(* IEC 61131-3 sources: daoli-st-library/DL_Device (part 5) *)

(* ---- FB_DL_RotaryAirlockCtrl.st ---- *)
(*==============================================================================
 * 组件名称 (Component)  : FB_DL_RotaryAirlockCtrl
 * 所属子库 (Sublibrary) : DL_Device
 * 当前版本 (Version)    : 1.0.2
 * 兼容性   (Platform)   : CODESYS 3.5 / TwinCAT 3 / 汇川 InoProShop / Machine Expert
 *                         仅依赖 Standard.library（TON / R_TRIG），零厂商方言
 * 来源标签 (Source)     : roadmap-industry-pool（粉体新方向 · 星型卸料器驱动，clean-room）
 * 功能描述 (Function)   : 星型卸料器（旋转气密阀）转速-料位联动驱动：
 *                         ① 料位联锁——高料位禁启（卡料风险），料位信号失效按
 *                            禁启（安全侧）；
 *                         ② 运行频率/转速给定（0..fFreqMax 钳位）；
 *                         ③ 电流失速判据——电流高于限值 AND 转速低于限值同拍
 *                            持续 tStallConfirm 确认窗 -> 停机 + 故障锁存；
 *                         ④ 反转点动解卡出口——仅停机态可用，受故障锁存闸拦截。
 * 范式次源 (Paradigm)   : 命令-反馈范式参照 I_DL_MotorDriver（CmdStart/CmdStop/
 *                         bRunning/bFault 契约），本件以引脚形式落地，不实现接口、
 *                         不引用接口方法（R31 家族纪律：只借范式不借实现）。
 * 高危区声明 (R31)      : 反转点动相与正转运行相为互斥高危区——两状态机分支互斥
 *                         由 CASE 结构保证（eJogRev 分支不产出任何正转输出，
 *                         eRunning / eStartPend 分支不产出反转输出），正反转输出
 *                         在统一出口再做一次 AND NOT 硬闸双保险。
 * 配比约束 (R100)       : tMinRun > tStallConfirm（最小运行窗必须宽于失速确认窗，
 *                         否则启动暂态电流尖峰会在转速未稳时被误判为失速）。
 * 边界与语义披露 (Boundary disclosure) :
 *   1) 料位联锁只禁启不停机：高料位 / 信号失效仅拒绝新的启动请求，运行中的
 *      卸料器不停（工艺侧决定），判据与码位按「拒启事件」承载。
 *   2) 电流 / 转速反馈非有限时失速判据挂起（不能拿垃圾信号判失速），但运行中
 *      反馈非有限本身升级为保护停机（故障级 030A，锁存至复位沿 + 信号恢复）。
 *   3) 启停频次守卫（DolMotor 判据口径）：停机后 tMinOff 未满拒绝再启动；
 *      信息级承载，不停摆、不锁存。
 *   4) 失速锁存解除路径（R152 自证可达）：复位沿 AND 失速条件已消失
 *      （电流回落 OR 转速回升）。
 * 故障码表 (Error codes) :
 *   16#0003_0507 [故障级] 失速确认窗满：停机 + 锁存，点动解卡被闸拦截
 *                 反证：停机 + eFault 与组态故障态输出组合不同但成因不可区分
 *                 （组态错 / 失速 / 反馈失效三因，必须码位互异 R190）。
 *   16#0003_0508 [故障级] 料位信号失效（无效标志或非有限），按禁启（锁存）
 *                 反证：禁启与高料位拒启输出组合相同，成因必须独立码位。
 *   16#0003_0509 [故障级] 组态非法（确认窗 / 限值域 / 频率上限），已两级回退
 *                 反证：回退后驱动照常，码位是组态错误唯一可见出口。
 *   16#0003_050A [故障级] 运行中电流 / 转速反馈非有限，保护停机 + 锁存
 *                 反证：保护停机与失速停机状态输出相同，成因必须独立码位。
 *   16#0003_0407 [信息级] 高料位拒启（启动请求被料位联锁拒绝）
 *                 反证：拒启事件 bStartRefused 为单拍脉冲，无码则拒因
 *                 （料位 / 频次 / 故障锁存）不可区分。
 *   16#0003_0408 [信息级] 启停频次守卫拒启（最小停机窗未满）
 *                 反证：频次守卫拒启与高料位拒启同为拒启脉冲，拒因组合不可区分。
 * 码位总账 (Code ledger) : 16#0003_0507 / 0508 / 0509 / 050A 用 ｜ 16#0003_0407 / 0408 用
 * 依赖     (Depends)    : 无 DL_ 内部依赖；Standard.library: TON / R_TRIG
 * 红线自检 (Redline)    : R1 ✓ 零全局变量与 VAR_EXTERNAL ｜ R2 ✓ 零 %I/%Q 物理地址
 *                         R3 ✓ 纯 IEC 61131-3 ｜ R4 ✓ 非有限双判 / 除数无涉 / 域闸全枚举
 *                         R5 ✓ 全变量中英双语同行注释 ｜ R6 ✓ 五态 ENUM + CASE + ELSE 兜底
 *                         R7 ✓ 四沿四计时主体最前部无条件刷新
 * 修订历史 (Revision)   :
 *   2026-11-22  v1.0.0  首版入库（R68 构建轮 · 批 2 · 目标 9）
 *   2026-11-22  v1.0.1  终审就地修①：组态锁存解除路径可达化（原 bCfgLatch 全文件零清零 -> 永久拒启）
 *   2026-11-22  v1.0.2  R69 点修⑥：正 / 反转出口改同拍派生（原 bJogRevOut 读上拍 bRunOut 反相，
 *                       反转首拍被上拍正转残值切断，滞后一拍；现两出口均由本拍状态派生，
 *                       交叉互斥在同一拍内完成）
 *============================================================================*)

(*-----------------------------------------------------------------------------
 * 枚举: E_DL_AirlockState（归属 DL_Device，与 FB_DL_RotaryAirlockCtrl 同文件）
 *----------------------------------------------------------------------------*)
TYPE E_DL_AirlockState :
(
    eIdle      := 0,    // 停机：可受理解卡点动 / Stopped, jog available
    eStartPend := 10,   // 启动命令已发，待运行反馈 / Start issued, awaiting run feedback
    eRunning   := 20,   // 运行反馈确认 / Running confirmed by feedback
    eJogRev    := 30,   // 反转点动解卡中（与正转互斥高危区）/ Reverse jog, exclusive with forward
    eFault     := 99    // 故障锁存：一切输出切断 / Fault latched, all outputs cut
);
END_TYPE

(*==============================================================================
 * 功能块: FB_DL_RotaryAirlockCtrl
 * 调用约定: 每个扫描周期无条件调用一次。
 *============================================================================*)
FUNCTION_BLOCK FB_DL_RotaryAirlockCtrl
VAR_INPUT
    bStartCmd       : BOOL;                  // 启动命令（电平）/ Start command, level
    bStopCmd        : BOOL;                  // 停止命令（电平，优先于启动）/ Stop command, level, priority
    bJogRevCmd      : BOOL;                  // 反转点动命令（电平，仅停机态有效）/ Reverse jog command, stopped only
    bRunFb          : BOOL;                  // 运行反馈（接触器 / 速度）/ Run feedback
    fLevelPct       : REAL;                  // 料位 [%] / Level [%]
    bLevelValid     : BOOL := TRUE;          // 料位信号有效标志 / Level signal valid flag
    fLevelHighLim   : REAL := 80.0;          // 高料位禁启阈 [%] / High level start-forbid threshold
    fFreqSet        : REAL := 25.0;          // 运行频率给定 [Hz] / Run frequency setpoint [Hz]
    fFreqMax        : REAL := 50.0;          // 频率上限 [Hz] / Frequency ceiling [Hz]
    fCurrent        : REAL;                  // 电机电流 [A] / Motor current [A]
    fSpeedFb        : REAL;                  // 转速反馈 [rpm] / Speed feedback [rpm]
    fStallCurrentLim: REAL := 10.0;          // 失速电流阈 [A] / Stall current threshold [A]
    fStallSpeedLim  : REAL := 1.0;           // 失速转速阈 [rpm] / Stall speed threshold [rpm]
    tStallConfirm   : TIME := T#3S;          // 失速确认窗 [s] / Stall confirmation window [s]
    tMinRun         : TIME := T#10S;         // 最小运行窗 [s] / Minimum run window [s]
    tMinOff         : TIME := T#30S;         // 最小停机窗 [s] / Minimum off window [s]
    bReset          : BOOL;                  // 上升沿：清除失速 / 料位 / 反馈失效锁存 / Rising edge: clear latches
END_VAR
VAR_OUTPUT
    bRunOut      : BOOL;                     // 正转运行输出（含启动待反馈段）/ Forward run output
    fFreqOut     : REAL;                     // 生效频率输出 [Hz] / Effective frequency output [Hz]
    bJogRevOut   : BOOL;                     // 反转点动输出 / Reverse jog output
    bStallLatch  : BOOL;                     // 失速锁存 / Stall latched
    bLevelBad    : BOOL;                     // 料位信号失效锁存 / Level signal invalid latched
    bStartRefused: BOOL;                     // 启动请求被拒脉冲（单拍）/ Start refused pulse, single scan
    bError       : BOOL;                     // 故障标志（锁存类归并）/ Fault flag, latched class merged
    uErrorId     : UDINT;                    // 故障码，0 = 无故障 / Error code, 0 = none
    eState       : E_DL_AirlockState;        // 当前状态（供 HMI 诊断）/ Current state for HMI diagnosis
END_VAR
VAR
    fbTrigStart  : R_TRIG;                  // 启动命令沿检测实例 / Start command edge detector
    fbTrigStop   : R_TRIG;                  // 停止命令沿检测实例 / Stop command edge detector
    fbTrigReset  : R_TRIG;                  // 复位沿检测实例 / Reset edge detector
    tonStall     : TON;                     // 失速确认窗计时实例 / Stall confirmation timer
    tonMinRun    : TON;                     // 最小运行窗计时实例 / Minimum run timer
    tonMinOff    : TON;                     // 最小停机窗计时实例 / Minimum off timer
    eStateInt    : E_DL_AirlockState;       // 主状态机内部当前态 / Internal state machine state
    bStallCond   : BOOL;                    // 本拍失速判据成立（反馈有效口径）/ Stall condition this scan
    bSigBadRun   : BOOL;                    // 运行中电流 / 转速非有限 / Current or speed non-finite while running
    bLevelNonFin : BOOL;                    // 料位非有限 / Level non-finite
    bLevelBadInt : BOOL;                    // 料位失效锁存内部副本 / Internal level-invalid latch
    bStallInt    : BOOL;                    // 失速锁存内部副本 / Internal stall latch
    bStartPermit : BOOL;                    // 本拍启动许可（料位口径）/ Start permit this scan, level class
    bFreqGuardOk : BOOL;                    // 本拍频次守卫通过 / Frequency guard passed
    fFreqClamp   : REAL;                    // 钳位后给定频率 [Hz] / Clamped setpoint frequency
    bCfgBad      : BOOL;                    // 本拍组态非法 / Config illegal this scan
    bCfgLatch    : BOOL;                    // 组态故障锁存（复位沿清除）/ Config fault latch
    bRefusedT    : BOOL;                    // 拒启脉冲内部副本（单拍）/ Internal refused pulse copy
    bErrorInt    : BOOL;                    // 本拍故障置位累加（出口归并）/ Fault set accumulator
    bFirstScan   : BOOL := TRUE;            // 上电首扫标志 / First-scan flag
END_VAR
VAR CONSTANT
    DL_RA_FIN_LIM : REAL := 1.0E30;   // REAL 有限幅值判界 / REAL finiteness bound
END_VAR

(*------------------------------------------------------------------------------
 * 段 1｜无条件刷新区（红线 R7）：四沿三计时全部位于主体最前部
 *      Unconditional refresh: four edges and three timers at the very top
 *      tonStall 的 IN 为内部派生判据（R40 断输入口径），禁挂外部引脚原值
 *-----------------------------------------------------------------------------*)
fbTrigStart(CLK := bStartCmd);
fbTrigStop(CLK := bStopCmd);
fbTrigReset(CLK := bReset);

bSigBadRun := (fCurrent <> fCurrent) OR (ABS(fCurrent) >= DL_RA_FIN_LIM)
              OR (fSpeedFb <> fSpeedFb) OR (ABS(fSpeedFb) >= DL_RA_FIN_LIM);
bLevelNonFin := (fLevelPct <> fLevelPct) OR (ABS(fLevelPct) >= DL_RA_FIN_LIM);

bStallCond := (eStateInt = E_DL_AirlockState.eRunning)
              AND (NOT bSigBadRun)
              AND (fCurrent > fStallCurrentLim)
              AND (fSpeedFb < fStallSpeedLim);

tonStall(IN := bStallCond, PT := tStallConfirm);
tonMinRun(IN := (eStateInt = E_DL_AirlockState.eRunning), PT := tMinRun);
tonMinOff(IN := (eStateInt = E_DL_AirlockState.eIdle), PT := tMinOff);

(*------------------------------------------------------------------------------
 * 段 2｜上电首扫：状态与输出落安全侧
 *      First-scan init: state and outputs to the safe side
 *-----------------------------------------------------------------------------*)
IF bFirstScan THEN
    eStateInt := E_DL_AirlockState.eIdle;
    fFreqClamp := 0.0;
    bFirstScan := FALSE;
END_IF

(*------------------------------------------------------------------------------
 * 段 3｜每拍预清（FB32-1）：单拍标志，禁入锁存 / 快照
 *      Per-scan preset: single-scan flags only
 *-----------------------------------------------------------------------------*)
bErrorInt  := FALSE;
bRefusedT  := FALSE;

(*------------------------------------------------------------------------------
 * 段 4｜组态域闸（R151 全枚举：四限值 + 三窗）+ 两级回退（R117）
 *      Config gate over all limits and windows, with two-level fallback
 *-----------------------------------------------------------------------------*)
bCfgBad := (tStallConfirm <= T#0S) OR (tMinRun <= T#0S) OR (tMinOff <= tMinRun)
           OR (fLevelHighLim <= 0.0) OR (fLevelHighLim > 100.0) OR (fLevelHighLim <> fLevelHighLim)
           OR (fStallCurrentLim <= 0.0) OR (fStallCurrentLim <> fStallCurrentLim)
           OR (fStallSpeedLim < 0.0) OR (fStallSpeedLim <> fStallSpeedLim)
           OR (fFreqMax <= 0.0) OR (fFreqMax <> fFreqMax);

IF bCfgBad THEN
    bCfgLatch := TRUE;
    uErrorId  := 16#0003_0509;   // 故障级：组态非法 / Fault: config illegal
    bErrorInt := TRUE;
END_IF

(* 终审就地修 v1.0.1（R68）：解除路径（R152 自证可达）——复位沿 AND 组态非法条件
 * 全部消失即清锁存。原实现把锁存清零只写在 eFault 相分支，而组态闸置锁存后
 * 并不迁相至 eFault（只回 eIdle / 驻留），eFault 相不可达 -> 锁存永不可解，
 * 组件保护/监视功能一次性永久失效直至 PLC 重启（终审两式①）。
 * Clear path made provably reachable: reset edge with the illegal config gone. *)
IF fbTrigReset.Q AND (NOT bCfgBad) THEN
    bCfgLatch := FALSE;          // 锁存解除 / Latch cleared
    uErrorId  := 16#0000_0000;   // 码位随解除归零 / Code cleared with the latch
END_IF

(*------------------------------------------------------------------------------
 * 段 5｜锁存类判据：料位失效（禁启）与运行反馈失效（保护停机）
 *      Latched criteria: level invalid forbids start, bad run feedback trips
 *      解除路径（R152 自证）：复位沿 AND 对应信号已恢复有效
 *-----------------------------------------------------------------------------*)
IF (NOT bLevelValid) OR bLevelNonFin THEN
    bLevelBadInt := TRUE;        // 失效按禁启（安全侧），不停运行（规格明示）/ Forbid start only
END_IF

(* 料位失效锁存解除路径（R152 自证可达）：复位沿 AND 料位信号已恢复有效 *)
(* Level latch clear path: reset edge AND the level signal valid again *)
IF fbTrigReset.Q AND bLevelValid AND (NOT bLevelNonFin) THEN
    bLevelBadInt := FALSE;
END_IF

IF bLevelBadInt THEN
    uErrorId  := 16#0003_0508;   // 故障级：料位信号失效 / Fault: level signal invalid
    bErrorInt := TRUE;
END_IF

IF bSigBadRun AND (eStateInt = E_DL_AirlockState.eRunning) THEN
    bStallInt := TRUE;           // 反馈失效按保护停机口径锁存 / Bad feedback trips protectively
    uErrorId  := 16#0003_050A;
    bErrorInt := TRUE;
    eStateInt := E_DL_AirlockState.eFault;   // 锁存同步迁相（FB50-1④）/ Latch migrates phase
END_IF

(*------------------------------------------------------------------------------
 * 段 6｜启动许可与频次守卫（边界 B1/B3）
 *      Start permit and frequency guard
 *-----------------------------------------------------------------------------*)
bStartPermit := bLevelValid AND (NOT bLevelNonFin) AND (fLevelPct < fLevelHighLim);
bFreqGuardOk := tonMinOff.Q;

(*------------------------------------------------------------------------------
 * 段 7｜主状态机（红线 R6）：ENUM + CASE + ELSE 兜底
 *      Main state machine with the mandatory ELSE fallback
 *-----------------------------------------------------------------------------*)
CASE eStateInt OF

    E_DL_AirlockState.eIdle:
        (* 停机相收到停止沿：无对象，事件湮灭（无状态改写，此处仅注释声明） *)
        (* Stop edge while idle: nothing to stop, event dies, no state write *)
        IF bJogRevCmd AND (NOT bRunFb) AND (NOT bStallInt) AND (NOT bLevelBadInt)
              AND (NOT bCfgLatch) THEN
            (* 反转点动（互斥高危区 R31）：仅停机态 + 无反馈 + 无故障锁存 *)
            (* Reverse jog: stopped, no feedback, no latch; exclusive high-risk zone *)
            eStateInt := E_DL_AirlockState.eJogRev;
        ELSIF fbTrigStart.Q THEN
            IF bStallInt OR bLevelBadInt OR bCfgLatch THEN
                bRefusedT := TRUE;       // 故障锁存类拒启 / Refused by a latch
                IF bStallInt THEN
                    uErrorId := 16#0003_0507;
                END_IF
            ELSIF NOT bStartPermit THEN
                bRefusedT := TRUE;       // 高料位 / 料位失效拒启 / Refused by level interlock
                uErrorId  := 16#0003_0407;
            ELSIF NOT bFreqGuardOk THEN
                bRefusedT := TRUE;       // 频次守卫拒启 / Refused by frequency guard
                uErrorId  := 16#0003_0408;
            ELSE
                eStateInt := E_DL_AirlockState.eStartPend;   // 受理，待反馈 / Accepted, awaiting feedback
            END_IF
        END_IF

    E_DL_AirlockState.eStartPend:
        IF bStopCmd OR fbTrigStop.Q OR bCfgLatch THEN
            eStateInt := E_DL_AirlockState.eIdle;    // 撤回 / Withdrawn
        ELSIF bRunFb THEN
            eStateInt := E_DL_AirlockState.eRunning; // 反馈确认 / Feedback confirmed
        END_IF

    E_DL_AirlockState.eRunning:
        IF bStopCmd OR fbTrigStop.Q OR bCfgLatch OR bStallInt THEN
            eStateInt := E_DL_AirlockState.eIdle;    // 停机 / 失速保护停机 / Stop or stall trip
        END_IF

    E_DL_AirlockState.eJogRev:
        IF bStopCmd OR bCfgLatch OR bStallInt OR (NOT bJogRevCmd) THEN
            eStateInt := E_DL_AirlockState.eIdle;    // 点动释放即回停机 / Jog release returns to idle
        END_IF

    E_DL_AirlockState.eFault:
        IF fbTrigReset.Q AND (NOT bStallCond) AND bLevelValid AND (NOT bLevelNonFin)
           AND (NOT bSigBadRun) AND (NOT bCfgBad) THEN
            bStallInt    := FALSE;       // 解除路径自证可达（R152）/ Clear path reachable
            bLevelBadInt := FALSE;
            uErrorId     := 16#0000_0000;
            eStateInt    := E_DL_AirlockState.eIdle;
        END_IF

    ELSE
        (* 非法状态拦截：切断一切输出，迁兜底态 *)
        eStateInt := E_DL_AirlockState.eFault;
        uErrorId  := 16#0003_0509;
        bErrorInt := TRUE;

END_CASE;

(*------------------------------------------------------------------------------
 * 段 8｜失速到期消化：确认窗满 -> 停机 + 锁存（与正常推进不同源，R 历史教训）
 *      Stall expiry digestion: window full trips stop and latch
 *      拍 N 进入：tonStall.Q 首次为真；本拍行为：置锁存 + 迁 eIdle；
 *      拍 N+1 转出：eIdle 相受复位沿 + 条件恢复解除
 *-----------------------------------------------------------------------------*)
IF tonStall.Q THEN
    bStallInt := TRUE;           // 失速锁存 / Stall latched
    uErrorId  := 16#0003_0507;   // 故障级：失速 / Fault: stall
    bErrorInt := TRUE;
    eStateInt := E_DL_AirlockState.eFault;   // 锁存同步迁相：停机 + 禁点动 / Latch migrates phase
END_IF

(*------------------------------------------------------------------------------
 * 段 9｜输出单一出口（范式 P-05）：正反转互斥硬闸（双保险，R31 高危区）
 *      Single output exit: forward and reverse outputs mutually exclusive
 *      R69 点修⑥：两出口一律由**本拍**状态派生后交叉互斥，禁止互相引用上拍输出
 *      （原实现 bJogRevOut := TRUE AND (NOT bRunOut) 读的是上一扫描的 bRunOut，
 *      反转首拍被上拍正转残值切断，解卡点动实际延后一拍；高危区出口不得有拍延迟）。
 *      Both outputs derive from the current phase, then cross-mask inside the same scan.
 *-----------------------------------------------------------------------------*)
bRunOut    := (eStateInt = E_DL_AirlockState.eRunning) OR (eStateInt = E_DL_AirlockState.eStartPend);
bJogRevOut := (eStateInt = E_DL_AirlockState.eJogRev);
bJogRevOut := bJogRevOut AND (NOT bRunOut);   // 反转串同拍正转非（双保险）/ Reverse masked by the same-scan forward
bRunOut    := bRunOut AND (NOT bJogRevOut);   // 正转串同拍反转非（双保险）/ Forward masked by the same-scan reverse

IF fFreqSet <> fFreqSet THEN
    fFreqOut := 0.0;                         // 给定非有限：频率安全侧 0 / Non-finite setpoint: safe zero
ELSIF fFreqSet < 0.0 THEN
    fFreqOut := 0.0;                         // 负给定钳 0 / Negative clamped
ELSIF fFreqSet > fFreqMax THEN
    fFreqOut := fFreqMax;                    // 超上限钳位 / Over clamped
ELSE
    fFreqOut := fFreqSet;                    // 合法直通 / Valid pass-through
END_IF

IF bCfgBad AND (fFreqMax <= 0.0) THEN
    fFreqOut := 0.0;                         // 上限组态非法时频率安全侧 0（R127 解耦）/ Safe zero when ceiling illegal
END_IF

bStallLatch := bStallInt;
bLevelBad   := bLevelBadInt;
bStartRefused := bRefusedT;                  // 单拍脉冲统一出口 / Unified single-scan exit
bError      := bErrorInt OR (eStateInt = E_DL_AirlockState.eFault);
eState      := eStateInt;
END_FUNCTION_BLOCK

(* ---- FB_DL_SafetyMuteZone.st ---- *)
(*==============================================================================
 * 组件名称 (Component)  : FB_DL_SafetyMuteZone
 * 所属子库 (Sublibrary) : DL_Device
 * 当前版本 (Version)    : 1.0.0
 * 兼容性   (Platform)   : CODESYS 3.5+ / TwinCAT 3 / 汇川 InoProShop / 施耐德 Machine Expert
 *                         仅依赖 Standard.library（TON / R_TRIG / F_TRIG），
 *                         零厂商私有库
 * 功能描述 (Function)   : 静默区（Muting）顺序时序判据：光幕遮挡（bLightCurtain=
 *                         TRUE=被遮挡）期间， mute 传感器须按 1→2 顺序激活才
 *                         合法静默（bMuted=TRUE）；2 先于 1 激活 → 乱序故障
 *                         锁存 bMuteFault（规格指定，R189 锁存回放）；静默窗
 *                         tMuteMax 超时 → 强制撤销静默回待机并置信息码
 *                         eMuteTimeout。合法时序：eIdle →（sen1 激活沿 ∧ 遮挡）
 *                         → eS1 →（sen2 激活沿）→ eMuted →（双释放 ∧ 光幕
 *                         恢复）→ eIdle。
 *                         **本件不作安全认证声明：仅作工艺物流静默时序编排，
 *                         人身安全由认证安全回路（安全 PLC/安全继电器）保证，
 *                         本件输出不得作为唯一安全切断依据。**
 * 接口     (Interface)  : 输入 bMuteSen1 静默传感器 1（TRUE=被物料遮挡）、
 *                         bMuteSen2 静默传感器 2、bLightCurtain 光幕（TRUE=
 *                         被遮挡）、tMuteMax 静默窗上限、bReset 复位；输出
 *                         bMuted 静默有效、bMuteFault 乱序故障锁存、ePhase
 *                         相位出口、eErrCode 错误码、bError 故障标志。
 * 边界     (Boundary)   : ① **属主边界（写死）：本件只做静默时序判据，不切断
 *                         光幕回路、不接管安全认证**（头注释安全声明）。
 *                         ② 四态 CASE + ELSE 兜底（R6）；tonMuteMax IN 挂
 *                         相驻留本身（eS1 ∨ eMuted 均计时，覆盖静默全程，
 *                         R145 使能域覆盖）；三沿实例段 0 无条件调用（R7）。
 *                         ③ 乱序归因唯一：sen2 先激活沿（eIdle 相内）→
 *                         eMuteFault 锁存 + eErrCode=eOrderBad；光幕未遮挡
 *                         期间传感器激活不作乱序（无静默语境）。
 *                         ④ 静默窗覆盖 eS1 与 eMuted 两相全程；超时强制撤销
 *                         回 eIdle（安全侧：静默撤销 = 光幕判据恢复有效），
 *                         信息码 eMuteTimeout 不锁存 bMuteFault（撤销本身为
 *                         安全侧动作）。
 *                         ⑤ 故障锁存解除路径：bMuteFault 解除边 = 传感器全
 *                         释放 ∧ bReset 上升沿（可达，头注释声明，R188）。
 *                         ⑥ 零全局耦合（无 GVL / VAR_EXTERNAL / 物理地址）。
 * 分工声明 (Scope)      : 与 `FB_DL_ElMutingGantry` 分工：龙门式静默布置归那件、
 *                         双传感器顺序静默区归本件；与 `FB_DL_FilmSpliceCurtain`
 *                         分工：拼接光幕归那件。
 * 来源标签 (Source Tag) : 自研线（双传感器静默顺序判据为公开物流静默模式
 *                         clean-room，不作安全认证声明）
 * 码表     (Codes)      : 本件不占用任何全局数字码位。出口为 BOOL 组 +
 *                         ENUM 相位/错误码；数字码位待主控收口阶段统一派号。
 * 红线自检 (Redline)    : R1 ✓ 零 GVL/VAR_EXTERNAL ｜ R2 ✓ 零 %I/%Q/%M ｜ R3 ✓ 纯 IEC 61131-3
 *                         R4 ✓ 乱序锁存解除可达 + 超时强制撤销安全侧 ｜ R5 ✓ 声明逐行同行双语注释
 *                         R6 ✓ 四态 CASE 含 ELSE ｜ R7 ✓ 一 TON 三沿段 0 无条件刷新
 * 修订历史 (Revision)   : 2026-11-20  v1.0.0  R50 首版（批次 4 · 序号 17）
 * 验收向量 (Acceptance) : ① 光幕遮挡后 sen1 激活、100ms 后 sen2 激活 → eMuted、
 *                         bMuted=TRUE；② 双传感器释放 ∧ 光幕恢复 → eIdle、
 *                         bMuted=FALSE；③ eIdle 相内 sen2 先激活 → bMuteFault
 *                         锁存、eErrCode=eOrderBad；④ 静默持续 > tMuteMax
 *                         → 强制回 eIdle、eErrCode=eMuteTimeout、bMuted=FALSE。
 *==============================================================================*)

(*-----------------------------------------------------------------------------
 * 枚举: E_DL_SmzPhase（静默区相位，全库唯一属主本文件）
 *----------------------------------------------------------------------------*)
TYPE E_DL_SmzPhase :
(
    eIdle  := 0,   // 待机（无静默语境） / Idle, no muting context
    eS1    := 10,  // 传感器 1 已激活（合法序列第 1 步） / Sensor 1 active, legal step one
    eMuted := 20,  // 静默有效（双传感器激活） / Muted, both sensors active
    eFault := 90   // 乱序故障（等复位） / Order fault, awaiting reset
);
END_TYPE

(*-----------------------------------------------------------------------------
 * 枚举: E_DL_SmzErr（错误码；信息级不置 bError，故障级恒伴 bError=TRUE）
 *----------------------------------------------------------------------------*)
TYPE E_DL_SmzErr :
(
    eOk          := 0,   // 正常 / Normal
    eOrderBad    := 1,   // 故障级：传感器乱序（2 先于 1） / Fault: sensor order violation
    eCfgBad      := 2,   // 故障级：静默窗组态非法（<= T#0S） / Fault: mute window config illegal
    eMuteTimeout := 3    // 信息级：静默窗超时强制撤销 / Info: mute window timeout, forced revoke
);
END_TYPE

FUNCTION_BLOCK FB_DL_SafetyMuteZone
VAR_INPUT
    bMuteSen1    : BOOL := FALSE;     // 静默传感器 1（TRUE=被物料遮挡） [-] / Muting sensor 1, TRUE blocked
    bMuteSen2    : BOOL := FALSE;     // 静默传感器 2（TRUE=被物料遮挡） [-] / Muting sensor 2, TRUE blocked
    bLightCurtain: BOOL := FALSE;     // 光幕（TRUE=被遮挡，静默语境前提） [-] / Light curtain, TRUE blocked
    tMuteMax     : TIME := T#30S;     // 静默窗上限，域 > T#0S [ms] / Mute window ceiling
    bReset       : BOOL := FALSE;     // 复位（须传感器全释放后上升沿才清故障锁存） [-] / Reset, clears fault when sensors released
END_VAR
VAR_OUTPUT
    bMuted   : BOOL;                  // 静默有效指示（eMuted 相电平） [-] / Muted indicator
    bMuteFault: BOOL;                 // 乱序故障锁存（解除 = 全释放 ∧ 复位沿） [-] / Order fault latch
    ePhase   : E_DL_SmzPhase;         // 相位出口 [-] / Phase outlet
    eErrCode : E_DL_SmzErr;           // 错误码出口 / Error code outlet
    bError   : BOOL;                  // 故障标志（乱序或组态） [-] / Error flag
END_VAR
VAR
    _eState   : E_DL_SmzPhase := E_DL_SmzPhase.eIdle;   // 内部相（CASE 唯一写入目标） / Internal phase
    _bFault   : BOOL;                 // 乱序故障锁存位（解除路径见头注释⑤） / Latched order fault bit
    _bCfgBad  : BOOL;                 // 组态非法当拍量 [-] / Illegal configuration
    _bCfgLatch: BOOL;                 // 组态故障锁存位（解除沿 = 全释放 ∧ bReset 上升沿） / Latched config fault
    _bTimeout : BOOL;                 // 静默窗超时当拍量（信息级） [-] / Mute timeout this scan
    rtReset   : R_TRIG;               // 复位沿实例，段 0 无条件调用 / Reset edge instance
    rtSen1    : R_TRIG;               // 传感器 1 激活沿实例，段 0 无条件调用 / Sensor 1 rising edge instance
    rtSen2    : R_TRIG;               // 传感器 2 激活沿实例，段 0 无条件调用 / Sensor 2 rising edge instance
    tonMuteMax: TON;                  // 静默窗 TON，段 0 无条件调用（IN 挂静默两相驻留，R145） / Mute window TON
END_VAR

(* —— 段 0：组态闸 + 全部沿/定时器无条件周期刷新（R6/R7） —— *)
_bCfgBad := (tMuteMax <= T#0S);       // 静默窗域闸 / Window configuration gate
rtReset(CLK := bReset);               // 复位沿，每拍必调 / Reset edge, every scan
rtSen1(CLK := bMuteSen1);             // 传感器 1 激活沿，每拍必调 / Sen 1 edge, every scan
rtSen2(CLK := bMuteSen2);             // 传感器 2 激活沿，每拍必调 / Sen 2 edge, every scan
tonMuteMax(IN := (_eState = E_DL_SmzPhase.eS1) OR (_eState = E_DL_SmzPhase.eMuted),
           PT := tMuteMax);           // 静默窗（覆盖 eS1/eMuted 全程，出相自复位） / Mute window covers both phases

(* —— 段 1：复位沿（须传感器全释放才清锁存，安全侧前提） —— *)
IF rtReset.Q AND (NOT bMuteSen1) AND (NOT bMuteSen2) THEN
    _bFault := FALSE;                 // 清乱序锁存（可达解除路径，头注释⑤） / Clear order fault
    _bCfgLatch := FALSE;              // 清组态锁存 / Clear config latch
    _eState := E_DL_SmzPhase.eIdle;   // 回待机 / Back to idle
END_IF
IF _bCfgBad AND (NOT _bCfgLatch) THEN
    _bCfgLatch := TRUE;               // 组态锁存 / Latch config fault
END_IF

(* —— 段 2：静默窗超时强制撤销（信息级；先于 CASE，撤销语义优先） —— *)
_bTimeout := tonMuteMax.Q AND (NOT _bFault) AND (NOT _bCfgLatch);   // 超时当拍量 / Timeout this scan
IF _bTimeout THEN
    _eState := E_DL_SmzPhase.eIdle;   // 强制撤销回待机（安全侧：光幕判据恢复有效） / Forced revoke to idle
END_IF

(* —— 段 3：四态顺控（故障/组态期冻结推进） —— *)
IF (NOT _bFault) AND (NOT _bCfgLatch) THEN
    CASE _eState OF

    E_DL_SmzPhase.eIdle:
        IF rtSen2.Q AND bLightCurtain THEN
            _bFault := TRUE;          // 乱序：sen2 先于 sen1 激活（规格③，归因唯一） / Order violation: sen 2 first
            _eState := E_DL_SmzPhase.eFault;   // 入故障相 / Enter fault
        ELSIF rtSen1.Q AND bLightCurtain THEN
            _eState := E_DL_SmzPhase.eS1;   // 合法第 1 步 / Legal step one
        END_IF

    E_DL_SmzPhase.eS1:
        IF rtSen2.Q THEN
            _eState := E_DL_SmzPhase.eMuted;   // 合法第 2 步：双激活静默 / Legal step two: muted
        ELSIF NOT bMuteSen1 THEN
            _eState := E_DL_SmzPhase.eIdle;   // sen1 提前释放：序列中止回待机 / Sequence aborted to idle
        END_IF

    E_DL_SmzPhase.eMuted:
        IF (NOT bMuteSen1) AND (NOT bMuteSen2) AND (NOT bLightCurtain) THEN
            _eState := E_DL_SmzPhase.eIdle;   // 双释放 ∧ 光幕恢复：静默结束 / Both released, curtain clear: end mute
        END_IF

    E_DL_SmzPhase.eFault:
        ;                            // 故障相驻留（由复位沿迁出链处理） / Held by reset chain

    ELSE
        _bFault := TRUE;             // 非法相位兜底（R45 配对见段 5） / Illegal phase fallback
        _eState := E_DL_SmzPhase.eFault;   // 强拉故障相 / Force fault phase

    END_CASE
END_IF

(* —— 段 4：出口单点映射（名实双出口同源，R191） —— *)
bMuted := (_eState = E_DL_SmzPhase.eMuted) AND (NOT _bFault) AND (NOT _bCfgLatch)
          AND (NOT _bTimeout);       // 静默有效出口（超时拍强制撤销） / Muted outlet
bMuteFault := _bFault;               // 故障锁存出口 / Fault latch outlet
ePhase := _eState;                   // 相位出口 / Phase outlet
IF _bCfgLatch THEN
    bError := TRUE;                  // 故障标志（R45 配对） / Error flag
    eErrCode := E_DL_SmzErr.eCfgBad; // 组态级码 / Config fault code
ELSIF _bFault THEN
    bError := TRUE;                  // 故障标志（乱序级） / Error flag
    eErrCode := E_DL_SmzErr.eOrderBad;   // 乱序锁存回放码（R189） / Order fault replay
ELSE
    bError := FALSE;                 // 无故障级条件 / No fault
    IF _bTimeout THEN
        eErrCode := E_DL_SmzErr.eMuteTimeout;   // 信息级：超时撤销 / Info: timeout revoke
    ELSE
        eErrCode := E_DL_SmzErr.eOk;            // 正常 / Normal
    END_IF
END_IF

END_FUNCTION_BLOCK

(* ---- FB_DL_SensorSupplyMon.st ---- *)
(*==============================================================================
 * 组件名称 (Component)  : FB_DL_SensorSupplyMon
 * 所属子库 (Sublibrary) : DL_Device
 * 当前版本 (Version)    : 1.0.0
 * 兼容性   (Platform)   : CODESYS 3.5+ / TwinCAT 3 / 汇川 InoProShop / 施耐德 Machine Expert
 *                         仅依赖 Standard.library（TON / ABS），零厂商私有库
 * 功能描述 (Function)   : 传感器供电轨监视（8 通道共用诊断掩码）：对供电实测
 *                         fSupplyMv（mV）做 tWindow 窗口均值（自复位 TON 窗，
 *                         窗内累加样本、窗到结算一次），再对窗口均值做迟滞判限：
 *                         均值 < fLimLowMv 入欠压态、恢复须均值 > fLimHighMv
 *                         （fLimLowMv < fLimHighMv 迟滞带，防临界振荡）；输出
 *                         bSupplyOk 与逐通道诊断掩码 uChanMask（bit i = 通道 i
 *                         使能 ∧ 供电正常）。非有限输入当拍跳过累计并置信息码
 *                         eInputHold，结论（bSupplyOk/掩码）保持上次值不翻转。
 * 接口     (Interface)  : 输入 fSupplyMv 供电实测 [mV]、tWindow 均值窗（域 > T#0S）、
 *                         fLimLowMv 欠压进入阈 [mV]、fLimHighMv 欠压恢复阈 [mV]、
 *                         uChanEn 8 通道使能位图（bit i=通道 i 参与诊断）、bReset
 *                         复位；输出 bSupplyOk 供电正常、uChanMask 逐通道诊断
 *                         掩码、fMeanMv 最新窗口均值 [mV]、eErrCode 错误码、
 *                         bError 故障标志。
 * 边界     (Boundary)   : ① **属主边界（写死）：本件只判供电轨好坏并出掩码，
 *                         不切换备用电源、不接管通道级断线诊断**；通道断线
 *                         诊断归 `FB_DL_AnalogTransmitter`。
 *                         ② 窗口均值：tonWin 自复位窗（IN := NOT tonWin.Q，
 *                         R188），窗内 fSum/nCnt 累计；窗到（Q 沿）结算一次
 *                         fMean = fSum ÷ nCnt，nCnt=0（整窗无非有限外样本）
 *                         跳过结算保持旧均值并置信息码，结构性无除零。
 *                         ③ 迟滞判限只在窗结算拍评估一次；判限态 _bLow 锁存，
 *                         进入阈 fLimLowMv < 恢复阈 fLimHighMv 构成迟滞带。
 *                         ④ 非有限样本（R79 双判）不计入累计：fSum/nCnt 不被
 *                         污染，当拍置 eInputHold 信息码，bSupplyOk 与掩码
 *                         保持上次结论（规格指定）。
 *                         ⑤ 组态闸：tWindow <= T#0S、fLimLowMv <= 0、
 *                         fLimHighMv <= fLimLowMv → 锁存故障，输出钳安全侧
 *                         bSupplyOk=FALSE，解除沿 = bReset 上升沿（故障级码
 *                         配对 bError，R45）。
 *                         ⑥ 掩码 bit i = uChanEn.bit i ∧ bSupplyOk ∧ 非 故障：
 *                         通道使能与供电结论逐位合成，定长 8 无越界。
 *                         ⑦ 零全局耦合（无 GVL / VAR_EXTERNAL / 物理地址）。
 * 分工声明 (Scope)      : 与 `FB_DL_MovingAverage` 分工：通用滑动平均归那件、
 *                         供电窗口均值+迟滞判限归本件；与 `FB_DL_AxiolineDiagLatch`
 *                         分工：总线级诊断锁存归那件。
 * 来源标签 (Source Tag) : 自研线（窗口均值+迟滞判限为公开监视模式 clean-room）
 * 码表     (Codes)      : 本件不占用任何全局数字码位。出口为 BOOL 组 + WORD 掩码
 *                         + LREAL 均值 + ENUM 错误码；数字码位待主控收口阶段
 *                         统一派号。
 * 红线自检 (Redline)    : R1 ✓ 零 GVL/VAR_EXTERNAL ｜ R2 ✓ 零 %I/%Q/%M ｜ R3 ✓ 纯 IEC 61131-3
 *                         R4 ✓ 除零前置闸 + 迟滞带 + 非有限保持结论 + 组态锁存
 *                         ｜ R5 ✓ 声明逐行同行双语注释
 *                         R6 N/A（无 ENUM 状态机，迟滞锁存态） ｜ R7 ✓ 一 TON 一 R_TRIG 段 0 无条件刷新
 * 修订历史 (Revision)   : 2026-11-20  v1.0.0  R50 首版（批次 1 · 序号 3）
 * 验收向量 (Acceptance) : ① tWindow=1s，窗内 10 个样本全 24000 mV → 均值
 *                         24000.0，24000 > fLimHighMv(22800) → bSupplyOk=
 *                         TRUE，uChanMask=使能位图全量；② 下一窗均值 22000 mV：
 *                         22000 < fLimLowMv(21600) 不成立且 > 恢复阈，迟滞带内
 *                         结论保持 TRUE（防临界振荡）；③ 窗均值 21000 mV <
 *                         21600 → bSupplyOk=FALSE、掩码全 0；④ 样本含 NaN：
 *                         该样本跳过、eErrCode=eInputHold，结论不翻转。
 *==============================================================================*)

(*-----------------------------------------------------------------------------
 * 枚举: E_DL_SsmErr（错误码；信息级不置 bError，故障级恒伴 bError=TRUE）
 *----------------------------------------------------------------------------*)
TYPE E_DL_SsmErr :
(
    eOk        := 0,   // 正常 / Normal
    eCfgBad    := 1,   // 故障级：组态非法（窗/阈值域） / Fault: illegal configuration
    eInputHold := 2    // 信息级：非有限输入跳过累计，结论保持 / Info: non-finite sample skipped, conclusion held
);
END_TYPE

FUNCTION_BLOCK FB_DL_SensorSupplyMon
VAR_INPUT
    fSupplyMv  : LREAL := 24000.0;    // 供电轨实测 [mV] / Supply rail measurement [mV]
    tWindow    : TIME := T#1S;        // 均值窗时长，域 > T#0S [ms] / Averaging window duration
    fLimLowMv  : LREAL := 21600.0;    // 欠压进入阈（均值低于此判欠压），域 > 0 [mV] / Undervolt entry threshold
    fLimHighMv : LREAL := 22800.0;    // 欠压恢复阈（须大于进入阈构成迟滞带） [mV] / Undervolt release threshold
    uChanEn    : WORD := 16#00FF;     // 8 通道使能位图（bit i=通道 i 参与诊断） [-] / Channel enable bitmap
    bReset     : BOOL := FALSE;       // 复位，上升沿清组态故障锁存 [-] / Reset, rising edge clears cfg latch
END_VAR
VAR_OUTPUT
    bSupplyOk  : BOOL;                // 供电正常（迟滞判限结论） [-] / Supply OK, hysteresis verdict
    uChanMask  : WORD;                // 逐通道诊断掩码（bit i=使能 ∧ 供电正常） [-] / Per-channel diagnostic mask
    fMeanMv    : LREAL;               // 最新有效窗口均值 [mV] / Latest valid window mean
    eErrCode   : E_DL_SsmErr;         // 错误码出口 / Error code outlet
    bError     : BOOL;                // 故障标志（组态锁存） [-] / Error flag, latched
END_VAR
VAR
    _fSum     : LREAL := 0.0;         // 窗内样本累计 [mV] / In-window sample sum
    _nCnt     : UDINT := 0;           // 窗内有效样本计数 [个] / In-window valid sample count
    _fMean    : LREAL := 0.0;         // 窗口均值锁存（结算源） [mV] / Window mean latch
    _bLow     : BOOL := FALSE;        // 欠压判限锁存态（迟滞源） [-] / Undervolt latched state
    _bBad     : BOOL := FALSE;        // 供电坏当拍结论（!bSupplyOk 内部量） [-] / Supply-bad verdict internal
    _bNonFin  : BOOL;                 // 当拍样本非有限 [-] / Sample non-finite this scan
    _bCfgBad  : BOOL;                 // 组态非法当拍量 [-] / Illegal configuration this scan
    _bSkip    : BOOL;                 // 本窗发生非有限跳过 [-] / Non-finite skip occurred in window
    _bWinEdge : BOOL;                 // 窗结算当拍量（Q 沿） [-] / Window settlement edge
    _bErrLatch: BOOL;                 // 组态故障锁存位（解除沿 = bReset 上升沿） / Latched config fault
    i         : DINT;                 // 通道循环索引 / Channel loop index
    rtReset   : R_TRIG;               // 复位沿实例，段 0 无条件调用 / Reset edge instance
    ftWin     : F_TRIG;               // 窗下降沿实例（Q 到结算一次），段 0 无条件调用 / Window F_TRIG settlement instance
    tonWin    : TON;                  // 自复位均值窗，段 0 无条件调用（R188） / Self-resetting averaging window
END_VAR
VAR CONSTANT
    DL_SSM_NCHAN : DINT := 8;         // 通道定长 [路] / Fixed channel count
    DL_SSM_BIT0  : WORD := 1;         // bit0 基准掩码 [-] / Bit zero base mask
    DL_SSM_ZERO  : LREAL := 0.0;      // 非有限判零基准与安全侧值 [mV] / Non-finite zero base and safe value
    DL_SSM_UDMAX : UDINT := 4294967295;   // 计数饱和点（防回绕） [个] / Count saturation ceiling
END_VAR

(* —— 段 0：非有限判 + 组态闸 + 窗口/沿无条件刷新 —— *)
_bNonFin := (fSupplyMv <> fSupplyMv) OR ((fSupplyMv - fSupplyMv) <> DL_SSM_ZERO);   // 样本非有限（R79 双判） / Sample non-finite
_bCfgBad := (tWindow <= T#0S) OR (fLimLowMv <= DL_SSM_ZERO)
         OR (fLimHighMv <= fLimLowMv);             // 组态域闸（窗/下阈/迟滞带方向） / Configuration gate
rtReset(CLK := bReset);                            // 复位沿，每拍必调 / Reset edge, every scan
tonWin(IN := (NOT tonWin.Q) AND (NOT _bErrLatch), PT := tWindow);   // 自复位均值窗（故障期停窗，R188） / Self-reset window, halted on fault
ftWin(CLK := tonWin.Q);                            // 窗结算沿，每拍必调 / Window settlement edge, every scan

(* —— 段 1：复位沿与组态闸入锁存 —— *)
IF rtReset.Q THEN
    _bErrLatch := FALSE;                           // 清组态锁存（R188 声明：解除沿 = bReset 上升沿） / Clear cfg latch
END_IF
IF _bCfgBad AND (NOT _bErrLatch) THEN
    _bErrLatch := TRUE;                            // 锁存 / Latch
END_IF

(* —— 段 2：窗内样本累计（非有限跳过并置信息量；故障期不累计） —— *)
_bSkip := FALSE;                                   // 本窗跳过量预清 / Window skip preset
IF (NOT _bErrLatch) AND (NOT _bNonFin) THEN
    _fSum := _fSum + fSupplyMv;                    // 有效样本累计 / Valid sample accumulate
    IF _nCnt < DL_SSM_UDMAX THEN
        _nCnt := _nCnt + 1;                        // 计数防回绕递增 / Count increment with wrap guard
    END_IF
ELSIF (NOT _bErrLatch) AND _bNonFin THEN
    _bSkip := TRUE;                                // 非有限样本跳过（不污染累计） / Non-finite sample skipped
END_IF

(* —— 段 3：窗结算（Q 下降沿一次；nCnt=0 跳过结算保持旧均值，无除零） —— *)
_bWinEdge := ftWin.Q;                              // 结算沿捕获 / Settlement edge capture
IF _bWinEdge AND (NOT _bErrLatch) THEN
    IF _nCnt > 0 THEN
        _fMean := _fSum / UDINT_TO_LREAL(_nCnt);   // 窗口均值（分母计数已判正） / Window mean, denominator proven positive
        IF _fMean < fLimLowMv THEN
            _bLow := TRUE;                         // 低于进入阈：判欠压 / Below entry threshold: undervolt
        ELSIF _fMean > fLimHighMv THEN
            _bLow := FALSE;                        // 高于恢复阈：解除欠压（迟滞带内保持） / Above release threshold: clear
        END_IF
        _bBad := _bLow;                            // 判限态落坏结论 / Verdict from hysteresis state
    END_IF
    _fSum := 0.0;                                  // 窗累计清零（下一窗重计） / Reset window sum
    _nCnt := 0;                                    // 窗计数清零 / Reset window count
END_IF

(* —— 段 4：掩码合成（bit i = 使能 ∧ 供电正常 ∧ 非故障；故障安全侧全 0） —— *)
FOR i := 0 TO (DL_SSM_NCHAN - 1) DO
    IF (NOT _bErrLatch) AND (NOT _bBad)
       AND ((uChanEn AND SHL(DL_SSM_BIT0, i)) <> 0) THEN
        uChanMask := uChanMask OR SHL(DL_SSM_BIT0, i);   // 通道 i 诊断通过（i∈[0,7] 位宽内） / Channel i passes
    ELSE
        uChanMask := uChanMask AND (NOT SHL(DL_SSM_BIT0, i));   // 通道 i 不通过：清位（禁直接跳过） / Channel i fails: clear bit
    END_IF
END_FOR

(* —— 段 5：出口单点映射（名实双出口同源，R191） —— *)
IF _bErrLatch THEN
    bSupplyOk := FALSE;                            // 故障安全侧：判供电坏 / Fault safe side: supply bad
    bError := TRUE;                                // 故障标志（R45 配对） / Error flag
    eErrCode := E_DL_SsmErr.eCfgBad;               // 故障级码 / Fault code
ELSE
    bSupplyOk := NOT _bBad;                        // 供电结论出口 / Supply verdict outlet
    bError := FALSE;                               // 无故障级条件 / No fault this scan
    IF _bSkip THEN
        eErrCode := E_DL_SsmErr.eInputHold;        // 信息级：结论保持口径 / Info: conclusion held
    ELSE
        eErrCode := E_DL_SsmErr.eOk;               // 正常 / Normal
    END_IF
END_IF
fMeanMv := _fMean;                                 // 均值出口（无有效窗保持旧值） / Mean outlet, held if no valid window

END_FUNCTION_BLOCK

(* ---- FB_DL_SlitValveInterlock.st ---- *)
(*==============================================================================
 * 组件名称 (Component)  : FB_DL_SlitValveInterlock
 * 溯源说明 (Provenance): 道莅 clean-room 防御性实现（IEC 61131-3 纯净实现，闭源文档仅借语义，零代码行）
 * 所属子库 (Sublibrary) : DL_Device / ValveInterlock
 * 当前版本 (Version)    : 1.0.0
 * 兼容性   (Platform)   : CODESYS 3.5 / TwinCAT 3 / 汇川 InoProShop / 施耐德
 *                         Machine Expert；纯 IEC 61131-3（第 3 版），仅用
 *                         Standard.library 的 TON / LIMIT
 * 组件分类 (Category)   : 功能块（FUNCTION_BLOCK）· 真空闸阀互斥互锁
 * 功能一句话 (Summary)  : 真空腔体与大传片腔之间的闸阀互锁：真空度、大气侧门位、
 *                         机械臂退出三个条件同拍判据，任一不满足即拒绝开阀并
 *                         给出位掩码阻塞原因；开/关指令严格互斥、先清后置。
 *
 * 本件存在的意义 (Why this unit exists)
 *   库内只有 InterlockMatrix 的通用掩码，没有「门类」语义：不知道真空度是
 *   模拟量、不知道门位反馈会自相矛盾、也不知道电磁阀开/关两路必须互斥。
 *   半导体 EFEM 场景里这些是必备项——闸阀在大气侧门开着时打开，等于把
 *   整个真空腔瞬间放空并可能夹住机械臂。
 *
 * 保守侧纪律 (Conservative side, 三条写死)
 *   ① 门位反馈自相矛盾（两路同时为真）或两路皆假持续 tFbTimeout
 *      → 故障 033D，**一律按「门未关」处理**（保守侧）；
 *   ② 真空度为非有限值或 < 0 → 故障 033E，**按「真空不足」处理**
 *      （不假定真空已建立）；
 *   ③ 联锁不满足而仍有开阀请求 → 故障 033C + uBlockMask（HMI 直接显示位）。
 *
 * 位置反馈收窄声明 (Pin truth —— 必须读，否则会误判本件缺陷)
 *   引脚集内**没有闸阀本体位置反馈**。tFbTimeout 的语义因此被收窄为
 *   「指令已发出但无位置确认」的等待窗：窗内保持指令且处于 eOpening；
 *   窗满仍无反馈则接受指令已生效、进 eOpen，并置信息 0173 提示
 *   「无位置反馈确认」。**绝不因超时反转指令**（规格④：保持指令并提示）。
 *   这不是遗漏，而是本件引脚契约的边界；有本体反馈的机型应在外部把反馈
 *   串入 bAtmDoorClosed/Open 的判据链，或另立带反馈的变体件。
 *
 * 边界安全 (Boundary)
 *   - 开/关两路输出**互斥**：段 1 先把两路都置 FALSE，段 8 再按状态只置一路
 *     （R72 双路径，同拍双 TRUE 是电磁阀线圈烧毁根因）；
 *   - 失能 → eClosing（先关阀），bValveOpenCmd := FALSE；关到位确认后回 eIdle；
 *   - 三个 TON 实例在主体前部无条件刷新（R40），门位/开等待/关等待各一只，
 *     绝不跨相复用同一实例；
 *   - CASE 落 ELSE 置 033E 兜底并回 eFault（非法状态无专用码，按「真空/判定
 *     不可信」同族复用，R90 留档）。
 *
 * 错误码    : 16#0003_0172 联锁满足，已放行开阀——信息级，正常放行
 *             16#0003_0173 到位反馈超时（无位置确认），保持当前指令——信息级，不反转
 *             16#0003_033C 联锁不满足，拒绝开阀（配 uBlockMask）——故障级
 *             16#0003_033D 门位反馈自相矛盾或缺失，按门未关处理——故障级
 *             16#0003_033E 真空度非法（非有限/负值/阈值非法），按真空不足处理——故障级
 * 码位总账  : 16#0003_0172 用 / 16#0003_0173 用 ｜ 16#0003_033C 用 / 16#0003_033D 用 / 16#0003_033E 用
 * 状态机    : E_DL_SlitValveState（eIdle / eOpening / eOpen / eClosing / eInterlock / eFault），
 *             CASE 含 ELSE 兜底，ELSE 置 16#0003_033E 并回 eFault；失能无条件回 eClosing
 * 采样约定  : 每任务周期调用一次；等待窗由 tFbTimeout 给定，不读系统时钟
 * 依赖说明  : 仅 Standard.library；健康出口本件不使用 E_DL_Ne107Status（互锁是
 *             许可判定而非健康分级），故不引用契约件
 * 验收向量  : V1 真空 50 Pa、门关、臂退、请求开 → 放行，eErr = 0172，bValveOpenCmd = TRUE，
 *                uBlockMask = 0，bInterlockOk = TRUE
 *             V2 真空 50 Pa、门两路同时为真 → 033D，uBlockMask 含位 2，拒绝开阀（保守侧主向量）
 *             V3 真空 -5 Pa → 033E，uBlockMask 含位 1，拒绝开阀（不假定真空主向量）
 *             V4 真空 500 Pa（> 阈值 100）、请求开 → 033C，uBlockMask = 1
 *             V5 请求开、门未关 → 033C + uBlockMask = 2，两路输出均为 FALSE（互斥向量）
 *             V6 请求开 3 s 无位置确认 → eOpen，eErr = 0173，指令保持 TRUE（不反转主向量）
 *             V7 bEnable 落 → eClosing，bValveOpenCmd = FALSE，关到位后回 eIdle
 * 红线自检  : 全局变量声明零使用 / 外部变量访问零使用 / 物理地址零使用 ｜ 纯 IEC 61131-3 ｜ 无除法
 *             浮点只用大小比较 ｜ 无循环 ｜ 全变量双语同行注释 ｜ ENUM + CASE 含
 *             ELSE ｜ 三个 TON 在主体前部无条件刷新 ｜ 位掩码常量化，无魔法数
 * 修订历史  : 2026-11-16  v1.0.0  首版入库（R22 · 批 2 · 设备安全互斥）
 *============================================================================*)

(*-----------------------------------------------------------------------------
 * 枚举: E_DL_SlitValveState（归属本功能块，同文件发布，全库唯一定义）
 * 含义: 闸阀互锁的工作相位。0 起步长 10。
 *-----------------------------------------------------------------------------*)
TYPE E_DL_SlitValveState :
(
    eIdle      := 0,   // 待机：阀关闭、无请求 / Idle, valve closed, no request
    eOpening   := 10,  // 开启中：指令已发，等待位置确认窗 / Opening, command issued, waiting for the ack window
    eOpen      := 20,  // 已开：指令保持有效 / Open, the command is held active
    eClosing   := 30,  // 关闭中：关阀指令有效 / Closing, the close command is active
    eInterlock := 40,  // 联锁阻塞：拒绝开阀并给出掩码 / Interlock blocked, opening refused with a mask
    eFault     := 99   // 故障：门位矛盾、真空非法或非法状态 / Fault, contradictory door, illegal vacuum or illegal state
);
END_TYPE

FUNCTION_BLOCK FB_DL_SlitValveInterlock
VAR_INPUT
    bRequest        : BOOL;                    // 开闸阀请求 / slit valve open request
    bAtmDoorClosed  : BOOL;                    // 大气侧门「已关」反馈 / atmospheric door closed feedback
    bAtmDoorOpen    : BOOL;                    // 大气侧门「已开」反馈 / atmospheric door open feedback
    fChamberVac     : REAL;                    // 腔体真空度 [Pa]，越小越真空 / chamber vacuum [Pa], the smaller the deeper
    fVacThreshold   : REAL := 100.0;           // 允许开闸阀的真空阈值 [Pa]，须 > 0 / vacuum threshold allowing opening [Pa], must be > 0
    bArmRetracted   : BOOL;                    // 机械臂已退出腔体 / robot arm retracted from the chamber
    tFbTimeout      : TIME := T#3S;            // 位置确认等待窗 [ms] / position acknowledgement window [ms]
    bEnable         : BOOL;                    // 使能 / enable
END_VAR
VAR_OUTPUT
    bValveOpenCmd   : BOOL;                    // 开阀指令，与关阀指令互斥 / open command, mutually exclusive with close
    bValveCloseCmd  : BOOL;                    // 关阀指令，与开阀指令互斥 / close command, mutually exclusive with open
    bInterlockOk    : BOOL;                    // 联锁全部满足 / all interlock conditions satisfied
    uBlockMask      : WORD;                    // 阻塞原因位掩码：1 真空不足 / 2 门未关 / 4 臂未退 / 8 反馈超时
    eErr            : UDINT;                   // 错误码，0 表示无错 / error code, 0 means no error
    bError          : BOOL;                    // 故障级标志，仅故障级错误置位 / fault-class flag, set only on fault-level codes
    bValid          : BOOL;                    // 输出可用标志 / outputs usable flag
END_VAR
VAR
    fbDoorWatch     : TON;                     // 门位反馈无效持续计时，段 5 无条件刷新 [ms] / door feedback invalid timer
    fbOpenWatch     : TON;                     // 开阀位置确认等待窗，段 5 无条件刷新 [ms] / open acknowledgement window
    fbCloseWatch    : TON;                     // 关阀位置确认等待窗，段 5 无条件刷新 [ms] / close acknowledgement window
    _eState         : E_DL_SlitValveState := E_DL_SlitValveState.eIdle; // 当前相位 / current phase
    _bInit          : BOOL := FALSE;           // 首扫标志，初值 FALSE 取非判定 / first-scan flag, tested negated
    _bIllegal       : BOOL;                    // 非法状态标志 / illegal state flag
    _bVacValid      : BOOL;                    // 真空度数值可用 / vacuum value usable
    _bVacOk         : BOOL;                    // 真空达标 / vacuum deep enough
    _bDoorValid     : BOOL;                    // 门位反馈有效（恰好一路为真） / door feedback valid, exactly one channel true
    _bDoorBadTime   : BOOL;                    // 门位反馈持续无效 / door feedback invalid for the whole window
    _bArmOk         : BOOL;                    // 机械臂已退出 / arm retracted
    _bBlkVac        : BOOL;                    // 阻塞位：真空不足 / block bit, vacuum insufficient
    _bBlkDoor       : BOOL;                    // 阻塞位：门未关 / block bit, door not closed
    _bBlkArm        : BOOL;                    // 阻塞位：臂未退 / block bit, arm not retracted
    _bBlkFb         : BOOL;                    // 阻塞位：反馈超时 / block bit, feedback timeout
    _bAllOk         : BOOL;                    // 三联条件全部满足 / all three conditions satisfied
    _bDoorBreak     : BOOL;                    // 门位计时器断输入一拍 / door timer one-scan break
    _bOpenBreak     : BOOL;                    // 开等待计时器断输入一拍 / open timer one-scan break
    _bCloseBreak    : BOOL;                    // 关等待计时器断输入一拍 / close timer one-scan break
    _tFbUse         : TIME := T#3S;            // 生效等待窗 [ms]，已钳位 / effective window, clamped
    _bAckTimeout    : BOOL;                    // 本拍发生确认超时 / acknowledgement timeout this scan
END_VAR
VAR CONSTANT
    DL_VAL_LIM      : REAL := 1.0E30;          // 有限性判定的绝对值上限 [Pa] / finiteness ceiling [Pa]
    DL_VAC_MIN      : REAL := 0.0;             // 真空度物理下限 [Pa]，负值非法 / vacuum physical floor [Pa], negatives illegal
    DL_THR_MIN      : REAL := 0.0;             // 真空阈值下限 [Pa]，须严格大于 / threshold floor [Pa], strictly greater
    DL_WIN_MIN_MS   : DINT := 1;               // 等待窗下限 [ms] / window floor [ms]
    DL_WIN_MAX_MS   : DINT := 60000;           // 等待窗上限 [ms] / window ceiling [ms]
    DL_BLK_VAC      : WORD := 16#0001;         // 掩码位 1：真空不足 / mask bit one, vacuum insufficient
    DL_BLK_DOOR     : WORD := 16#0002;         // 掩码位 2：大气门未关 / mask bit two, atmospheric door not closed
    DL_BLK_ARM      : WORD := 16#0004;         // 掩码位 4：机械臂未退 / mask bit four, arm not retracted
    DL_BLK_FB       : WORD := 16#0008;         // 掩码位 8：反馈超时 / mask bit eight, feedback timeout
    DL_MASK_NONE    : WORD := 16#0000;         // 无阻塞 / no blocking
END_VAR

(*------------------------------------------------------------------------------
 * 段 1｜每拍预置：两路输出**先清后置**（R72，互斥的唯一保证手段）
 *      Every scan starts with both commands cleared, exclusivity is structural
 *-----------------------------------------------------------------------------*)
bValveOpenCmd  := FALSE;                       // 开阀指令先清 / open command cleared first
bValveCloseCmd := FALSE;                       // 关阀指令先清 / close command cleared first
bInterlockOk   := FALSE;                       // 联锁满足位预置 FALSE / interlock ok preset FALSE
uBlockMask     := DL_MASK_NONE;                // 掩码清零 / mask cleared
eErr           := 16#0000_0000;                // 错误码预置无错 / error code preset to none
bError         := FALSE;                       // 故障标志预置 FALSE / fault flag preset to FALSE
bValid         := FALSE;                       // 输出可用预置 FALSE / usable flag preset to FALSE
_bIllegal      := FALSE;                       // 非法状态标志预清零 / illegal state flag pre-cleared
_bVacValid     := FALSE;                       // 真空可用标志预清零 / vacuum usable pre-cleared
_bVacOk        := FALSE;                       // 真空达标标志预清零 / vacuum ok pre-cleared
_bDoorValid    := FALSE;                       // 门位有效标志预清零 / door valid pre-cleared
_bDoorBadTime  := FALSE;                       // 门位持续无效标志预清零 / door bad time pre-cleared
_bArmOk        := FALSE;                       // 臂退出标志预清零 / arm ok pre-cleared
_bBlkVac       := FALSE;                       // 真空阻塞位预清零 / vacuum block pre-cleared
_bBlkDoor      := FALSE;                       // 门阻塞位预清零 / door block pre-cleared
_bBlkArm       := FALSE;                       // 臂阻塞位预清零 / arm block pre-cleared
_bBlkFb        := FALSE;                       // 反馈阻塞位预清零 / feedback block pre-cleared
_bAllOk        := FALSE;                       // 全条件标志预清零 / all-ok pre-cleared
_bAckTimeout   := FALSE;                       // 确认超时标志预清零 / ack timeout pre-cleared

(*------------------------------------------------------------------------------
 * 段 2｜首扫初始化（阀位默认关闭：失电安全位）
 *      First-scan initialisation, the valve defaults closed
 *-----------------------------------------------------------------------------*)
IF NOT _bInit THEN
    _eState     := E_DL_SlitValveState.eIdle;  // 相位待机 / phase idle
    _bDoorBreak := TRUE;                       // 门位计时从零开始 / door timer starts from zero
    _bOpenBreak := TRUE;                       // 开等待计时从零开始 / open timer starts from zero
    _bCloseBreak := TRUE;                      // 关等待计时从零开始 / close timer starts from zero
    _bInit      := TRUE;                       // 首扫只做一次 / the first scan runs once
END_IF

(*------------------------------------------------------------------------------
 * 段 3｜真空度判定（非有限 / 负值 / 阈值非法 → 按「真空不足」处理）
 *      Vacuum evaluation, invalid values are treated as insufficient
 *-----------------------------------------------------------------------------*)
IF (fVacThreshold <> fVacThreshold) OR (ABS(fVacThreshold) > DL_VAL_LIM)
   OR (fVacThreshold <= DL_THR_MIN) THEN
    _bVacValid := FALSE;                       // 阈值非法：真空判定不可信 / illegal threshold, the vacuum test is untrustworthy
ELSE
    IF (fChamberVac < -DL_VAL_LIM) OR (fChamberVac > DL_VAL_LIM) THEN
        _bVacValid := FALSE;                   // 非有限值：不可用 / non-finite value
    ELSIF fChamberVac < DL_VAC_MIN THEN
        _bVacValid := FALSE;                   // 负压读数非法：不可用 / negative reading is illegal
    ELSE
        _bVacValid := TRUE;                    // 数值可用 / the value is usable
        _bVacOk    := (fChamberVac <= fVacThreshold); // 真空达标判据 [布尔] / deep enough test
    END_IF
END_IF
IF NOT _bVacValid THEN
    eErr := 16#0003_033E;                      // 故障级：真空度非法，按不足处理 / fault: illegal vacuum, treated as insufficient
    bError := TRUE;                            // 置故障标志 / raise the fault flag
    _bVacOk := FALSE;                          // 不假定真空（保守侧） / never assume vacuum
END_IF

(*------------------------------------------------------------------------------
 * 段 4｜门位反馈有效性（恰好一路为真才算有效；矛盾与缺失都按门未关）
 *      Door feedback validity, exactly one channel must be true
 *-----------------------------------------------------------------------------*)
_bDoorValid := (bAtmDoorClosed OR bAtmDoorOpen) AND (NOT (bAtmDoorClosed AND bAtmDoorOpen));

(*------------------------------------------------------------------------------
 * 段 5｜三个计时器无条件刷新（R40：CASE 之外每拍必调，各相各一只实例）
 *      Three timers refreshed unconditionally outside the CASE, one instance each
 *-----------------------------------------------------------------------------*)
_tFbUse := tFbTimeout;                         // 等待窗直取引脚 [ms] / window taken from the pin
IF TIME_TO_DINT(_tFbUse) < DL_WIN_MIN_MS THEN
    _tFbUse := DINT_TO_TIME(DL_WIN_MIN_MS);    // 下限钳位（1 ms），防零窗每拍超时 / clamped to the floor
END_IF
IF TIME_TO_DINT(_tFbUse) > DL_WIN_MAX_MS THEN
    _tFbUse := DINT_TO_TIME(DL_WIN_MAX_MS);    // 上限钳位（60 s） / clamped to the ceiling
END_IF

fbDoorWatch(IN := (NOT _bDoorValid) AND (NOT _bDoorBreak), PT := _tFbUse); // 门位持续无效计时
_bDoorBreak := FALSE;                          // 断输入拍在调用后自清 / break self-cleared after the call
_bDoorBadTime := fbDoorWatch.Q;                // 持续无效达窗口 / invalid for the whole window

fbOpenWatch(IN := (_eState = E_DL_SlitValveState.eOpening) AND (NOT _bOpenBreak), PT := _tFbUse); // 开阀确认等待窗
_bOpenBreak := FALSE;                          // 断输入拍在调用后自清 / break self-cleared

fbCloseWatch(IN := (_eState = E_DL_SlitValveState.eClosing) AND (NOT _bCloseBreak), PT := _tFbUse); // 关阀确认等待窗
_bCloseBreak := FALSE;                         // 断输入拍在调用后自清 / break self-cleared

(*------------------------------------------------------------------------------
 * 段 6｜联锁判据与掩码拼装（三条全部写进掩码，便于现场一次定位）
 *      Interlock criteria and mask assembly, every criterion lands in the mask
 *-----------------------------------------------------------------------------*)
_bArmOk := bArmRetracted;                      // 机械臂退出判据 / arm retracted test
_bBlkVac  := NOT _bVacOk;                      // 真空不足（含数值非法） / vacuum insufficient, invalid included
_bBlkDoor := NOT (bAtmDoorClosed AND (NOT bAtmDoorOpen)); // 门未关（含矛盾与缺失） / door not closed, contradictions included
_bBlkArm  := NOT _bArmOk;                      // 臂未退 / arm not retracted
_bBlkFb   := _bDoorBadTime;                    // 反馈持续无效 / feedback invalid for the whole window

IF _bBlkVac THEN
    uBlockMask := uBlockMask OR DL_BLK_VAC;    // 置真空不足位 / set the vacuum bit
END_IF
IF _bBlkDoor THEN
    uBlockMask := uBlockMask OR DL_BLK_DOOR;   // 置门未关位 / set the door bit
END_IF
IF _bBlkArm THEN
    uBlockMask := uBlockMask OR DL_BLK_ARM;    // 置臂未退位 / set the arm bit
END_IF
IF _bBlkFb THEN
    uBlockMask := uBlockMask OR DL_BLK_FB;     // 置反馈超时位 / set the feedback bit
END_IF

_bAllOk := (_bVacOk AND (NOT _bBlkDoor) AND _bArmOk AND (NOT _bBlkFb)); // 三联条件全部满足
bInterlockOk := _bAllOk;                       // 联锁满足出口 / interlock ok outlet

(*------------------------------------------------------------------------------
 * 段 7｜相位机（只做迁移；两路指令在段 8 按状态置位）
 *      Phase machine, transitions only, the commands are set in segment eight
 *-----------------------------------------------------------------------------*)
CASE _eState OF

    E_DL_SlitValveState.eIdle:                 // 待机：有请求且联锁满足才允许开
        IF (NOT _bDoorValid AND _bDoorBadTime) THEN
            _eState := E_DL_SlitValveState.eFault; // 门位持续无效，转故障 / door feedback persistently invalid
            eErr    := 16#0003_033D;           // 故障级：门位反馈矛盾或缺失 / fault: contradictory or missing door feedback
            bError  := TRUE;                   // 置故障标志 / raise the fault flag
        ELSIF bEnable AND bRequest THEN
            IF _bAllOk THEN
                _eState := E_DL_SlitValveState.eOpening; // 联锁满足，放行开阀 / interlock ok, allow opening
                _bOpenBreak := TRUE;           // 开等待窗从零开始 / the open window starts from zero
                eErr    := 16#0003_0172;       // 信息级：已放行开阀 / informational: opening released
            ELSE
                _eState := E_DL_SlitValveState.eInterlock; // 联锁不满足，转阻塞 / blocked
                eErr    := 16#0003_033C;       // 故障级：拒绝开阀 / fault: opening refused
                bError  := TRUE;               // 置故障标志 / raise the fault flag
            END_IF
        END_IF

    E_DL_SlitValveState.eOpening:              // 开启中：等待确认窗；窗满接受指令已生效
        IF (NOT _bDoorValid AND _bDoorBadTime) THEN
            _eState := E_DL_SlitValveState.eFault; // 门位持续无效，转故障 / door feedback persistently invalid
            eErr    := 16#0003_033D;           // 故障级：门位反馈矛盾或缺失 / fault: contradictory or missing door feedback
            bError  := TRUE;                   // 置故障标志 / raise the fault flag
        ELSIF (NOT bEnable) OR (NOT bRequest) THEN
            _eState := E_DL_SlitValveState.eClosing; // 请求撤销或失能：先关阀 / request dropped or disabled, close first
            _bCloseBreak := TRUE;              // 关等待窗从零开始 / the close window starts from zero
        ELSIF NOT _bAllOk THEN
            _eState := E_DL_SlitValveState.eClosing; // 条件转差：先关阀（安全侧） / conditions degraded, close
            _bCloseBreak := TRUE;              // 关等待窗从零开始 / the close window starts from zero
        ELSIF fbOpenWatch.Q THEN
            _eState := E_DL_SlitValveState.eOpen; // 窗满无反馈：接受指令已生效 / window elapsed, treat the command as effective
            _bAckTimeout := TRUE;              // 标记确认超时 / flag the acknowledgement timeout
            eErr    := 16#0003_0173;           // 信息级：无位置确认，保持指令 / informational: no position confirmation, command held
        END_IF

    E_DL_SlitValveState.eOpen:                 // 已开：条件转差或请求撤销即关
        IF (NOT _bDoorValid AND _bDoorBadTime) THEN
            _eState := E_DL_SlitValveState.eFault; // 门位持续无效，转故障 / door feedback persistently invalid
            eErr    := 16#0003_033D;           // 故障级：门位反馈矛盾或缺失 / fault: contradictory or missing door feedback
            bError  := TRUE;                   // 置故障标志 / raise the fault flag
        ELSIF (NOT bEnable) OR (NOT bRequest) OR (NOT _bAllOk) THEN
            _eState := E_DL_SlitValveState.eClosing; // 任一条件撤销：关阀 / any condition lost, close
            _bCloseBreak := TRUE;              // 关等待窗从零开始 / the close window starts from zero
        END_IF

    E_DL_SlitValveState.eClosing:              // 关闭中：关到位（窗满）后回待机
        IF _bAllOk AND bEnable AND bRequest AND fbCloseWatch.Q THEN
            _eState := E_DL_SlitValveState.eOpening; // 关闭窗满且条件满足：重新开 / close window elapsed, reopen
            _bOpenBreak := TRUE;               // 开等待窗从零开始 / the open window starts from zero
            eErr    := 16#0003_0172;           // 信息级：已放行开阀 / informational: opening released
        ELSIF fbCloseWatch.Q THEN
            _eState := E_DL_SlitValveState.eIdle; // 关到位，回待机 / closed, back to idle
        END_IF

    E_DL_SlitValveState.eInterlock:            // 联锁阻塞：条件恢复且仍有请求才放行
        IF NOT bEnable THEN
            _eState := E_DL_SlitValveState.eIdle; // 失能回待机（保持关阀） / disabled, back to idle, keep closed
        ELSIF NOT bRequest THEN
            _eState := E_DL_SlitValveState.eIdle; // 请求撤销回待机 / request dropped
        ELSIF _bAllOk THEN
            _eState := E_DL_SlitValveState.eOpening; // 条件恢复，放行开阀 / conditions restored
            _bOpenBreak := TRUE;               // 开等待窗从零开始 / the open window starts from zero
            eErr    := 16#0003_0172;           // 信息级：已放行开阀 / informational: opening released
        ELSE
            eErr    := 16#0003_033C;           // 故障级：仍然拒绝开阀 / fault: still refused
            bError  := TRUE;                   // 置故障标志 / raise the fault flag
        END_IF

    E_DL_SlitValveState.eFault:                // 故障：门位恢复有效且真空可用才回待机
        IF _bDoorValid AND _bVacValid THEN
            _eState := E_DL_SlitValveState.eIdle; // 原因消失，回待机 / cause cleared, back to idle
        END_IF

    ELSE
        _bIllegal := TRUE;                     // 标记非法状态 / flag the illegal state
        _eState   := E_DL_SlitValveState.eFault; // 回故障态 / back to the fault state
        eErr      := 16#0003_033E;             // 兜底复用：判定不可信（R90 不加码） / fallback reuse: untrustworthy evaluation
        bError    := TRUE;                     // 置故障标志 / raise the fault flag
END_CASE

(*------------------------------------------------------------------------------
 * 段 8｜指令输出（严格互斥：段 1 已全清，此处最多置一路）
 *      Command outputs, strictly exclusive, at most one is set here
 *-----------------------------------------------------------------------------*)
CASE _eState OF
    E_DL_SlitValveState.eOpening:              // 开启中：只置开阀 / opening, only the open command
        bValveOpenCmd := TRUE;                 // 开阀指令 / open command
    E_DL_SlitValveState.eOpen:                 // 已开：保持开阀指令 / open, hold the open command
        bValveOpenCmd := TRUE;                 // 开阀指令 / open command
    E_DL_SlitValveState.eClosing:              // 关闭中：只置关阀 / closing, only the close command
        bValveCloseCmd := TRUE;                // 关阀指令 / close command
    E_DL_SlitValveState.eInterlock:            // 阻塞：只置关阀（保守侧，绝不留开阀） / blocked, close only
        bValveCloseCmd := TRUE;                // 关阀指令 / close command
    E_DL_SlitValveState.eFault:                // 故障：只置关阀 / fault, close only
        bValveCloseCmd := TRUE;                // 关阀指令 / close command
    ELSE
        bValveCloseCmd := FALSE;               // 待机与非法状态：两路指令均为 FALSE（阀由弹簧/自保持停在失电安全位） / idle, no command asserted
END_CASE

(*------------------------------------------------------------------------------
 * 段 9｜出口与可用性仲裁（码位优先级：故障级 > 信息级）
 *      Exit and usability arbitration
 *-----------------------------------------------------------------------------*)
IF _bAckTimeout AND (NOT bError) AND (eErr = 16#0000_0000) THEN
    eErr := 16#0003_0173;                      // 信息级：确认超时（不反转指令） / informational: ack timeout
END_IF

IF bError OR _bIllegal THEN
    bValid := FALSE;                           // 故障级或非法状态：输出不可用 / fault or illegal state: outputs unusable
ELSIF NOT bEnable THEN
    bValid := FALSE;                           // 失能：输出不可用 / disabled: unusable
ELSE
    bValid := TRUE;                            // 输出可用 / outputs usable
END_IF

END_FUNCTION_BLOCK

(* ---- FB_DL_StatusWordSegDecoder.st ---- *)
(*==============================================================================
 * 组件名称 (Component)  : FB_DL_StatusWordSegDecoder
 * 所属子库 (Sublibrary) : DL_Device
 * 当前版本 (Version)    : 1.0.0
 * 组件分类 (Category)   : 功能块（FUNCTION_BLOCK）· 设备状态字 · 段表驱动解码
 * 兼容性   (Platform)   : CODESYS 3.5 / TwinCAT 3 / 汇川 InoProShop / Schneider
 *                         Machine Expert；仅 SHL / SHR 位运算与标准类型
 * 功能描述 (Function)   : 用一张段描述表（最多 16 段，每段含位偏移、位宽与
 *                         名称）把设备状态字一次性解码成右对齐的值数组，并在
 *                         同一拍给出越界、重叠、段数三类组态诊断与段状态位。
 *                         替代「每字段调用一次单段提取」的碎片写法：一次调用
 *                         拿全部字段，且组态错误在投运首日即被拦下。
 * 双宽域声明 (Width)    : 入口统一为 64 位宽字，DWORD 调用方把高位补零即可。
 *                         宽度是参数域而非语义差异，故不拆 32 位与 64 位两块。
 * 边界声明 (Boundary)   : FC_DL_BitGet 取单个位；FB_DL_UnpackWordToBits 拆固定
 *                         十六位；FC_DL_BitFieldExtract 取单段；FC_DL_WordBitPack
 *                         做单段打包。四者均为「单点」件，本块是本族唯一的
 *                         「组态级」件：段表驱动的 N 段批量解码加段间重叠诊断，
 *                         且位段提取在本块内自写，不调用上述任何单段件。
 * 掩码构造纪律 (Mask)   : 宽度等于 64 时直接取全 1 常量，**不**做 64 位移位
 *                         （对 64 位字移位 64 是未定义行为，跨平台结果不一致）。
 *                         其余宽度按「低位连续 1 左移偏移」两步构造，宽度与
 *                         偏移都在段级校验通过后才参与移位。
 * 重叠语义 (Overlap)    : 用 64 位占位掩码逐段求与，非零即重叠。拒绝模式
 *                         （bRejectOnOverlap 为真）下后到段整段作废；覆盖模式
 *                         下后到段生效（取后段值），占位掩码同步合并。两种模式
 *                         都置段状态位与信息级码，组态问题不会被静默吞掉。
 * 开源溯源 (Origin)     : lgf-bitlogic / rockwell-aoi / plcnext-community。参考
 *                         公开位逻辑功能库与设备 AOI 的段描述参数组织方式
 *                         （偏移、宽度、名称三元组）以及状态字解码的功能分类，
 *                         只借参数组织与分类，位序、掩码构造、重叠算法、枚举、
 *                         状态机、码位与全部实现 100% 自有，clean-room 实现，
 *                         不构成衍生作品。
 * 依赖     (Depends)    : 无 DL_ 内部依赖；仅 Standard.library 的 SHL / SHR
 * 故障码表 (Error codes):
 *   16#0003_0142【信息级】段间重叠（拒绝模式下该段作废，覆盖模式下取后段）
 *   16#0003_0143【信息级】段越界已拒绝（宽度为零、宽度超字宽、偏移加宽超字宽）
 *   16#0003_0144【信息级】段数越界已钳位（小于 1 或大于 16）
 *   16#0003_0302【故障级】段表整体非法（无任何段可用）或非法状态兜底
 * 码位占用 (Slot)       : 信息级 0142 / 0143 / 0144；故障级 0302。
 *                         全部落在 R11 本件分配块内，无跨块借用。
 * 写入点次序 (Write order) :
 *   ① uSegStatusMask ：段解码段逐段置位，本拍起点清零，全拍只增不覆写
 *   ② auValue        ：段解码段逐段写，未定义段与作废段一律写 0
 *   ③ ePhase         ：状态机段为唯一位移点，复位分支只回待机
 *   ④ uErrorId       ：输出段单一优先级链（0302 优于 0142 优于 0143 优于 0144）
 * 验收向量 (Acceptance) :
 *   V1 单段跨半字节：字 16#1234、段（偏移 4、宽度 8）→ 值 16#23 = 35
 *   V2 双段：段（4,8）与段（8,8）→ 值 35 与 16#12 = 18
 *   V3 重叠：段（0,8）与段（4,8）、拒绝模式 → 状态掩码 16#0003、有效段 1、
 *      码 16#0003_0142
 *   V4 越界：段（60,8）→ 该段值为 0、状态位置位、码 16#0003_0143，其余段不受影响
 *   V5 六十四位特例：段（0,64）且字全 1 → 值 16#FFFF_FFFF，全程无 64 位移位
 * 红线自检 (Redline)    : R1 零全局变量表与外部变量引用 ｜ R2 零物理地址直写
 *                         R3 纯 IEC 61131-3 ｜ R4 段级边界先校验后移位，无除零
 *                         R5 全变量中英双语同行注释 ｜ R6 ENUM 加 CASE 加 ELSE
 *                         R7 R_TRIG 在 CASE 之外无条件刷新
 *                         R8 信息级码 0142 至 0144 不置组态故障位
 * 修订历史 (Revision)   :
 *   2026-11-15  v1.0.0  首版落盘（Round 11 · 泳道 B · 位段批量解码开组）
 *============================================================================*)

(*------------------------------------------------------------------------------
 * 结构体: ST_DL_BitSeg（单段描述：偏移、宽度、名称）
 *         One segment descriptor, offset, width and a readable name
 *-----------------------------------------------------------------------------*)
TYPE ST_DL_BitSeg :
STRUCT
    nOffset : USINT;        // 段起始位偏移 [位]，有效域 0 到 63 / Segment start bit offset, zero to sixty-three
    nWidth  : USINT;        // 段位宽 [位]，有效域 1 到 64 / Segment width in bits, one to sixty-four
    sName   : STRING[16];   // 段名称 [文本]，供 HMI 显示与排故定位 / Segment name for the HMI and for troubleshooting
END_STRUCT
END_TYPE

(*------------------------------------------------------------------------------
 * 结构体: ST_DL_BitSegTable（段描述表容器，由调用方组态并持有）
 *         Segment descriptor table container, configured and owned by the caller
 *-----------------------------------------------------------------------------*)
TYPE ST_DL_BitSegTable :
STRUCT
    aSeg      : ARRAY[1..16] OF ST_DL_BitSeg;  // 段描述数组，十六段上限 [段] / Segment descriptor array, sixteen entries maximum
    nReserved : INT;                           // 预留字段，保持结构体对齐惯例 [整数] / Reserved field keeping the library struct convention
END_STRUCT
END_TYPE

(*------------------------------------------------------------------------------
 * 枚举: E_DL_SegDecodePhase（本块相位，归属本功能块并同文件发布）
 *       Phase enumeration owned by this block and published in the same file
 *-----------------------------------------------------------------------------*)
TYPE E_DL_SegDecodePhase :
(
    eIdle   := 0,   // 待机：未使能，值数组清零 / Idle, value array cleared
    eDecode := 10,  // 解码：逐拍重解，值随源字刷新 / Decoding, re-evaluated every cycle
    eReject := 20,  // 拒绝：整表无可用段，组态故障，需改表并复位 / Rejected, no usable segment, fix the table and reset
    eFault  := 99   // 故障：非法相位兜底，需复位退出 / Fault, illegal phase fallback, needs a reset
);
END_TYPE

(*==============================================================================
 * 逐拍推演 (Cycle-by-cycle trace)：
 *   场景 A 两段正常（段一偏移 4 宽 8，段二偏移 8 宽 8，字 16#1234）
 *     段解码段：段一掩码为高位连续八位左移四位，取值 16#23 得 35，占位合并；
 *          段二掩码不与占位相交，取值 16#12 得 18，占位合并；有效段计数为 2
 *     状态机段：eDecode 自保持；输出段有效段 2、段状态掩码 0、码 0
 *   场景 B 重叠且拒绝模式（段一 0 宽 8，段二 4 宽 8）
 *     段一正常取值并占位；段二掩码与占位相交，置段状态位两位，段二作废；
 *          有效段计数为 1；输出段码 16#0003_0142，组态故障位保持假
 *   场景 C 越界（段三偏移 60 宽 8）
 *     段级校验先做：偏移加宽 68 超过 64，直接拒绝，不参与移位、不参与占位；
 *          该段值写 0，其余段照常解码，码 16#0003_0143
 *   场景 D 整表不可用（唯一段宽度为 0）
 *     有效段计数为 0 → eReject、组态故障位为真、码 16#0003_0302；
 *          改表后有效段计数回到 1，复位上升沿退回待机，下一拍重入解码
 *   场景 E 六十四位特例（段一 0 宽 64，字全 1）
 *     宽度等于字宽直接取全 1 常量，不做移位；取值低 32 位为 16#FFFF_FFFF
 *============================================================================*)

(*==============================================================================
 * 状态迁移表 (State transition table)：
 *   当前相位   迁移条件                          目标相位   伴随动作
 *   eIdle      使能为真                          eDecode    值数组在解码段刷新
 *   eDecode    有效段数大于等于 1                eDecode    自保持，逐拍重解
 *   eDecode    有效段数为 0 且请求段数大于等于 1 eReject    组态故障位为真
 *   eDecode    使能为假                          eIdle      值数组清零
 *   eReject    使能为假                          eIdle      值数组清零
 *   eReject    复位沿且有效段数大于等于 1        eIdle      表已修正，回待机重入
 *   eFault     复位沿                            eIdle      非法相位标记清除
 *   其他值     任意                              eFault     码归入 0302
 *   说明：eReject 不自动恢复——组态问题必须人工确认后复位，避免「表错但
 *   偶发可用」时反复跳变；而 eDecode 允许逐拍重解，源字变化立即反映到值数组。
 *============================================================================*)

(*==============================================================================
 * 掩码构造对照表 (Mask construction)：
 *   段位宽   掩码构造方式                     注意事项
 *   1       单比特基准左移偏移                最常用，等价取单个标志位
 *   2 到 31 低位连续一左移后整体左移偏移      两步走，先造宽度再定位
 *   32      低位连续一左移后整体左移偏移      低半字取值，高位被自然丢弃
 *   33 到 63 同上，仍在 64 位字内合法          宽度与偏移之和不得超 64
 *   64      直接取全 1 常量                    禁对 64 位字移位 64，属未定义行为
 *   0       直接判越界拒绝                     宽度为零无物理意义
 *   说明：宽度大于 64 或偏移加宽超 64 一律在段级校验拦下，绝不进入移位分支；
 *   这是「先校验后运算」纪律的具体落点，与浮点先判零再除法同源。
 *============================================================================*)

(*==============================================================================
 * 重叠模式对照表 (Overlap policy)：
 *   项目           拒绝模式（真）              覆盖模式（假）
 *   后到段取值     写 0，整段作废              取后段值，后写者生效
 *   占位掩码       不合并                      合并，后续段继续判重叠
 *   有效段计数     不计该段                    计入
 *   段状态位       置位                        置位（重叠事实不变）
 *   信息级码       0142                        0142
 *   适用场合       字段定义严格、不允许歧义     上级字含兼容旧定义的冗余字段
 *   说明：两种模式都置段状态位与信息级码，重叠绝不会被静默吞掉；选择哪一种
 *   由调用方按设备手册的字段定义决定，本块不替现场做语义判断。
 *============================================================================*)

(*==============================================================================
 * 段表组态投运检查清单 (Commissioning checklist)：
 *   ① 段数：请求段数不超过十六，且与段表实际填写段数一致（多填的段不解码）
 *   ② 单调性：段偏移无需递增，但重叠必须是有意为之，否则投运首日就会看到 0142
 *   ③ 满宽段：宽度等于 64 的段只允许存在一段，且偏移必须为 0
 *   ④ 名称：段名建议写设备手册原文缩写，排故时与手册逐条对照
 *   ⑤ 字节序：本块只做位序解码，多字节字段的高低字节交换请在 IO 映射层完成，
 *      不要在段表里用两个半字节段去拼一个整字，那样会触发重叠诊断
 *   说明：以上五条是现场投运阶段最常见的组态错误来源，本块把它们转成段状态
 *   位与信息级码，让问题在第一次上电时就暴露，而不是等到三个月后偶发停机。
 *============================================================================*)

FUNCTION_BLOCK FB_DL_StatusWordSegDecoder
VAR_INPUT
    bEnable           : BOOL;                       // 使能，FALSE 时值数组清零 [-] / Enable, clears the value array on FALSE
    bReset            : BOOL;                       // 清组态诊断，上升沿有效 [-] / Clears the configuration diagnostics on a rising edge
    uWord             : LWORD;                      // 被解码状态字，六十四位宽 [位串] / Source status word, sixty-four bits wide
    nSegCount         : INT;                        // 有效段数 [段]，有效域 1 到 16 / Valid segment count, one to sixteen
    bRejectOnOverlap  : BOOL;                       // 重叠策略，真为整段拒绝，假为后段覆盖 [-] / Overlap policy, reject the segment or let the later one win
END_VAR
VAR_OUTPUT
    auValue           : ARRAY[1..16] OF UDINT;      // 各段解码值，右对齐，未定义段为 0 [值] / Decoded value per segment, right aligned, zero for unused
    nValidCount       : INT;                        // 实际成功解码的段数 [段] / Segment count successfully decoded
    uSegStatusMask    : WORD;                       // 段状态位：置位表示该段越界或重叠被拒 [位串] / Segment status bits, set when rejected
    eState            : E_DL_SegDecodePhase;        // 主状态机当前相位 [-] / Current phase of the main state machine
    bConfigFault      : BOOL;                       // 段表组态故障（整表无可用段）[-] / Segment table configuration fault
    uErrorId          : UDINT;                      // 事件码，0 表示无事件 [代码] / Event code, zero means none
END_VAR
VAR_IN_OUT
    stSegs            : ST_DL_BitSegTable;          // 段描述表，块内只读，禁止就地改写 [-] / Segment descriptor table, read only inside this block
END_VAR
VAR
    fbTrigReset       : R_TRIG;                     // 复位沿检测，CASE 之外无条件刷新 [-] / Reset edge detector, refreshed outside the CASE
    bInit             : BOOL := FALSE;              // 首扫标志，初值 FALSE，判据 NOT bInit [-] / First-scan flag initialised FALSE
    ePhase            : E_DL_SegDecodePhase := E_DL_SegDecodePhase.eIdle;  // 内部相位，对外经 eState 输出 / Internal phase, exported as eState
    nSegClamped       : INT;                        // 钳位后的段数 [段]，0 到 16 / Clamped segment count, zero to sixteen
    bSegCntClamped    : BOOL;                       // 段数越界被钳位的标记 [-] / Flag, segment count was clamped
    bSegCntEmpty      : BOOL;                       // 段数小于一的标记 [-] / Flag, segment count below one
    nWidthUse         : INT;                        // 当前段位宽 [位] / Width of the current segment
    nOffsetUse        : INT;                        // 当前段位偏移 [位] / Bit offset of the current segment
    uSegMask          : LWORD;                      // 当前段掩码 [位串] / Mask of the current segment
    uOccupy           : LWORD;                      // 已占位掩码，重叠检测用 [位串] / Occupied bit mask used for overlap detection
    bSegBad           : BOOL;                       // 当前段越界标记 [-] / Flag, current segment is out of range
    bSegDup           : BOOL;                       // 当前段重叠标记 [-] / Flag, current segment overlaps a previous one
    bAnyOut           : BOOL;                       // 本拍存在越界段 [-] / Flag, at least one segment is out of range
    bAnyOverlap       : BOOL;                       // 本拍存在重叠段 [-] / Flag, at least one segment overlaps
    bStateIllegal     : BOOL;                       // 非法相位被兜底捕获 [-] / Flag, an illegal phase was captured
    i                 : INT;                        // 段遍历索引 [1..16] / Segment loop index
END_VAR
VAR CONSTANT
    DL_SEG_MAX        : INT := 16;                  // 段数上限 [段] / Maximum segment count
    DL_WORD_BITS      : INT := 64;                  // 位宽常量 [位] / Word width in bits
    DL_MASK64_ALL     : LWORD := 16#FFFF_FFFF_FFFF_FFFF;  // 六十四位全 1 掩码 [位串] / All ones mask for the full width
    DL_MASK64_ONE     : LWORD := 16#0000_0000_0000_0001;  // 六十四位单比特基准 [位串] / Single bit reference of the full width
    DL_MASK64_NONE    : LWORD := 16#0000_0000_0000_0000;  // 六十四位全 0 掩码 [位串] / All zeros mask
    DL_MASK_ONE       : WORD := 16#0001;            // 段状态位单比特基准 [位串] / Single bit reference for the status mask
    DL_SEG_MIN        : INT := 1;                   // 段数下限 [段] / Minimum segment count
    DL_WIDTH_MIN      : INT := 1;                   // 段宽下限 [位] / Minimum segment width
END_VAR

(*------------------------------------------------------------------------------
 * 段 1｜沿检测无条件刷新（R7 红线）
 *      Edge detection refreshed unconditionally
 *-----------------------------------------------------------------------------*)
fbTrigReset(CLK := bReset);

(*------------------------------------------------------------------------------
 * 段 2｜首扫初始化（R19 唯一合法范式）
 *      First-scan initialisation with the canonical R19 pattern
 *-----------------------------------------------------------------------------*)
IF NOT bInit THEN
    FOR i := 1 TO DL_SEG_MAX DO
        auValue[i] := 0;                 // 值数组初值确定，HMI 不显示随机数
    END_FOR
    nValidCount     := 0;
    uSegStatusMask  := 16#0000;
    ePhase          := E_DL_SegDecodePhase.eIdle;
    eState          := E_DL_SegDecodePhase.eIdle;
    bConfigFault    := FALSE;
    bStateIllegal   := FALSE;
    uErrorId        := 16#0000_0000;
    bInit           := TRUE;             // 首扫只做一次
END_IF

(*------------------------------------------------------------------------------
 * 段 3｜段数钳位（小于一整体不动作，大于上限钳位到十六）
 *      Segment count clamping, below one does nothing, above sixteen clamped
 *-----------------------------------------------------------------------------*)
bSegCntClamped := FALSE;
bSegCntEmpty   := FALSE;
IF nSegCount < DL_SEG_MIN THEN
    nSegClamped   := 0;                  // 无有效段：整体不动作
    bSegCntEmpty  := TRUE;
ELSIF nSegCount > DL_SEG_MAX THEN
    nSegClamped   := DL_SEG_MAX;         // 超上限钳位
    bSegCntClamped := TRUE;
ELSE
    nSegClamped := nSegCount;
END_IF

(*------------------------------------------------------------------------------
 * 段 4｜段解码（段级校验先于移位；重叠用占位掩码求与判定）
 *      Segment decoding, validation before shifting, overlap by occupy mask
 *      位段提取在本块内自写，不调用任何单段提取件，保证泳道内零跨依赖
 *      每段处理分三步，顺序不可颠倒：
 *        第一步 校验：宽度小于一、宽度超字宽、偏移加宽超字宽，任一成立即拒绝，
 *               该段不参与移位、不参与占位，仅置段状态位与越界标记
 *        第二步 造掩码：满宽特例走全 1 常量，其余走「连续一左移」两步构造
 *        第三步 取值与占位：取值写值数组；拒绝模式下重叠段写 0 且不合并占位，
 *               覆盖模式下取值并合并占位，有效段计数同步加一
 *-----------------------------------------------------------------------------*)
uOccupy        := DL_MASK64_NONE;
uSegStatusMask := 16#0000;
nValidCount    := 0;
bAnyOut        := FALSE;
bAnyOverlap    := FALSE;
FOR i := 1 TO DL_SEG_MAX DO
    auValue[i] := 0;                                     // 未定义段与作废段一律为 0
END_FOR

IF bEnable AND (ePhase <> E_DL_SegDecodePhase.eFault) THEN
    FOR i := 1 TO nSegClamped DO
        nWidthUse  := USINT_TO_INT(stSegs.aSeg[i].nWidth);
        nOffsetUse := USINT_TO_INT(stSegs.aSeg[i].nOffset);
        bSegBad    := FALSE;
        bSegDup    := FALSE;

        IF (nWidthUse < DL_WIDTH_MIN)
           OR (nWidthUse > DL_WORD_BITS)
           OR ((nOffsetUse + nWidthUse) > DL_WORD_BITS) THEN
            bSegBad := TRUE;                             // 段级越界：先拒绝，后不参与移位
        END_IF

        IF bSegBad THEN
            uSegStatusMask := uSegStatusMask OR SHL(DL_MASK_ONE, i - 1);
            bAnyOut        := TRUE;
        ELSE
            IF nWidthUse >= DL_WORD_BITS THEN
                uSegMask := DL_MASK64_ALL;               // 满宽特例：禁 64 位移位
            ELSE
                uSegMask := SHL(DL_MASK64_ONE, nWidthUse) - DL_MASK64_ONE;
                uSegMask := SHL(uSegMask, nOffsetUse);   // 低位连续一左移到位
            END_IF

            IF (uOccupy AND uSegMask) <> DL_MASK64_NONE THEN
                uSegStatusMask := uSegStatusMask OR SHL(DL_MASK_ONE, i - 1);
                bAnyOverlap    := TRUE;
                bSegDup        := TRUE;
            END_IF

            IF bSegDup AND bRejectOnOverlap THEN
                auValue[i] := 0;                         // 拒绝模式：后到段整段作废
            ELSE
                auValue[i] := LWORD_TO_UDINT(SHR(uWord AND uSegMask, nOffsetUse));
                uOccupy    := uOccupy OR uSegMask;       // 覆盖模式：占位合并，后段生效
                nValidCount := nValidCount + 1;
            END_IF
        END_IF
    END_FOR
END_IF

(*------------------------------------------------------------------------------
 * 段 5｜主状态机（ENUM 加 CASE，含 ELSE 兜底；每成员均有对应标签）
 *      Main state machine, one label per enumeration member plus a fallback
 *-----------------------------------------------------------------------------*)
CASE ePhase OF
    E_DL_SegDecodePhase.eIdle:
        IF bEnable THEN
            ePhase := E_DL_SegDecodePhase.eDecode;       // 使能即进入逐拍重解
        END_IF

    E_DL_SegDecodePhase.eDecode:
        IF NOT bEnable THEN
            ePhase := E_DL_SegDecodePhase.eIdle;
        ELSIF (nValidCount = 0) AND (nSegClamped >= DL_SEG_MIN) THEN
            ePhase := E_DL_SegDecodePhase.eReject;       // 整表无可用段：组态故障
        END_IF

    E_DL_SegDecodePhase.eReject:
        IF NOT bEnable THEN
            ePhase := E_DL_SegDecodePhase.eIdle;
        ELSIF fbTrigReset.Q AND (nValidCount >= DL_SEG_MIN) THEN
            ePhase := E_DL_SegDecodePhase.eIdle;         // 表已修正且复位：退回待机重入
        END_IF

    E_DL_SegDecodePhase.eFault:
        IF fbTrigReset.Q THEN
            ePhase        := E_DL_SegDecodePhase.eIdle;  // 只有复位可退出兜底故障
            bStateIllegal := FALSE;
        END_IF

    ELSE
        ePhase        := E_DL_SegDecodePhase.eFault;     // 非法值兜底
        bStateIllegal := TRUE;
END_CASE

(*------------------------------------------------------------------------------
 * 段 6｜输出归并与码位定级（单一优先级链，全拍只写一次 uErrorId）
 *      Output merge and single-priority error code resolution
 *-----------------------------------------------------------------------------*)
IF NOT bEnable THEN
    FOR i := 1 TO DL_SEG_MAX DO
        auValue[i] := 0;                                 // 未使能一律清零，避免陈旧值
    END_FOR
    nValidCount := 0;
    uSegStatusMask := 16#0000;
END_IF

bConfigFault := bStateIllegal
                OR (bEnable AND (nSegClamped >= DL_SEG_MIN) AND (nValidCount = 0));

IF bConfigFault THEN
    uErrorId := 16#0003_0302;                            // 优先级一：整表非法
ELSIF bAnyOverlap THEN
    uErrorId := 16#0003_0142;                            // 信息级：段间重叠
ELSIF bAnyOut THEN
    uErrorId := 16#0003_0143;                            // 信息级：段越界已拒绝
ELSIF bSegCntClamped OR bSegCntEmpty THEN
    uErrorId := 16#0003_0144;                            // 信息级：段数越界已钳位
ELSE
    uErrorId := 16#0000_0000;
END_IF

eState := ePhase;                                        // 相位每拍重写，供 HMI 诊断
END_FUNCTION_BLOCK
